FUNCTION "FRK_ModelRoot" : Int
{ S7_Optimized_Access := 'TRUE' }
VERSION : 0.1
VAR_INPUT
    Scope : String;
END_VAR
BEGIN
    #FRK_ModelRoot := 0;
    IF #Scope = 'StationA' THEN #FRK_ModelRoot := 1; RETURN; END_IF;
    IF #Scope = 'StationB' THEN #FRK_ModelRoot := 2; RETURN; END_IF;
END_FUNCTION
// Core model identities and cloned configuration are one owned catalog domain.
// Native UMAC/recipe CSV cannot replace its typed, root-scoped admission rules.
FUNCTION "FRK_ModelCodeValid" : Bool
{ S7_Optimized_Access := 'TRUE' }
VERSION : 0.1
VAR_INPUT Code : String; END_VAR
VAR_TEMP Index : Int; Value : Byte; END_VAR
BEGIN
    #FRK_ModelCodeValid := FALSE;
    IF LEN(#Code) < 1 OR LEN(#Code) > 64 THEN RETURN; END_IF;
    FOR #Index := 1 TO LEN(#Code) DO
        #Value := CHAR_TO_BYTE(#Code[#Index]);
        IF #Value < BYTE#32 OR #Value > BYTE#126 THEN RETURN; END_IF;
    END_FOR;
    #FRK_ModelCodeValid := TRUE;
END_FUNCTION

FUNCTION "FRK_ModelCrc" : DWord
{ S7_Optimized_Access := 'TRUE' }
VERSION : 0.1
VAR_IN_OUT Catalog : "FRK_ModelCatalog"; END_VAR
VAR_TEMP Work : DWord; Index : Int; Character : Int; Size : Int; Text : String[80]; END_VAR
BEGIN
    #Work := "FRK_CrcNumber"(Previous := DWORD#16#FFFFFFFF, Value := UINT_TO_UDINT(#Catalog.SchemaVersion));
    #Size := LEN(#Catalog.Scope);
    #Work := "FRK_CrcNumber"(Previous := #Work, Value := INT_TO_UDINT(#Size));
    FOR #Character := 1 TO #Size DO #Work := "FRK_CrcByte"(Previous := #Work, Value := CHAR_TO_BYTE(#Catalog.Scope[#Character])); END_FOR;
    #Work := "FRK_CrcNumber"(Previous := #Work, Value := INT_TO_UDINT(#Catalog.Capacity));
    #Work := "FRK_CrcNumber"(Previous := #Work, Value := INT_TO_UDINT(#Catalog.Count));
    #Work := "FRK_CrcNumber"(Previous := #Work, Value := #Catalog.Generation);
    FOR #Index := 1 TO 3 DO
        #Text := #Catalog.Codes[#Index]; #Size := LEN(#Text);
        #Work := "FRK_CrcNumber"(Previous := #Work, Value := INT_TO_UDINT(#Size));
        FOR #Character := 1 TO #Size DO #Work := "FRK_CrcByte"(Previous := #Work, Value := CHAR_TO_BYTE(#Text[#Character])); END_FOR;
    END_FOR;
    #FRK_ModelCrc := NOT #Work;
END_FUNCTION

FUNCTION "FRK_ModelValid" : Bool
{ S7_Optimized_Access := 'TRUE' }
VERSION : 0.1
VAR_INPUT RootIndex : Int; END_VAR
VAR_IN_OUT Catalog : "FRK_ModelCatalog"; END_VAR
VAR_TEMP Index : Int; Other : Int; END_VAR
BEGIN
    #FRK_ModelValid := FALSE;
    IF #RootIndex < 1 OR #RootIndex > 2 OR "FRK_ModelRoot"(Scope := #Catalog.Scope) <> #RootIndex THEN RETURN; END_IF;
    IF #Catalog.SchemaVersion <> 1 OR #Catalog.Generation = 0 OR #Catalog.Capacity <> 3
        OR #Catalog.Count < 2 OR #Catalog.Count > 3 THEN RETURN; END_IF;
    IF #Catalog.Codes[1] <> 'MODEL_A' OR #Catalog.Codes[2] <> 'MODEL_B' THEN RETURN; END_IF;
    FOR #Index := 1 TO #Catalog.Count DO
        IF NOT "FRK_ModelCodeValid"(Code := #Catalog.Codes[#Index]) THEN RETURN; END_IF;
        FOR #Other := 1 TO #Index - 1 DO
            IF #Catalog.Codes[#Index] = #Catalog.Codes[#Other] THEN RETURN; END_IF;
        END_FOR;
    END_FOR;
    FOR #Index := #Catalog.Count + 1 TO 3 DO
        IF #Catalog.Codes[#Index] <> '' THEN RETURN; END_IF;
    END_FOR;
    #FRK_ModelValid := #Catalog.Checksum = "FRK_ModelCrc"(Catalog := #Catalog);
END_FUNCTION

FUNCTION "FRK_ModelVirgin" : Bool
{ S7_Optimized_Access := 'TRUE' }
VERSION : 0.1
VAR_IN_OUT Catalog : "FRK_ModelCatalog"; END_VAR
VAR_TEMP Index : Int; END_VAR
BEGIN
    #FRK_ModelVirgin := FALSE;
    IF #Catalog.SchemaVersion <> 0 OR #Catalog.Scope <> '' OR #Catalog.Capacity <> 0 OR #Catalog.Count <> 0
        OR #Catalog.Generation <> 0 OR #Catalog.Checksum <> DWORD#0 THEN RETURN; END_IF;
    FOR #Index := 1 TO 3 DO IF #Catalog.Codes[#Index] <> '' THEN RETURN; END_IF; END_FOR;
    #FRK_ModelVirgin := TRUE;
END_FUNCTION

FUNCTION "FRK_ModelKnown" : Bool
{ S7_Optimized_Access := 'TRUE' }
VERSION : 0.1
VAR_INPUT RootIndex : Int; Code : String; END_VAR
VAR_TEMP Index : Int; END_VAR
BEGIN
    #FRK_ModelKnown := FALSE;
    IF #RootIndex < 1 OR #RootIndex > 2 OR #Code = '' THEN RETURN; END_IF;
    IF "FRK_ModelStore".Rows[#RootIndex].Count < 2 OR "FRK_ModelStore".Rows[#RootIndex].Count > 3 THEN RETURN; END_IF;
    FOR #Index := 1 TO "FRK_ModelStore".Rows[#RootIndex].Count DO
        IF "FRK_ModelStore".Rows[#RootIndex].Codes[#Index] = #Code THEN #FRK_ModelKnown := TRUE; RETURN; END_IF;
    END_FOR;
END_FUNCTION
FUNCTION "FRK_ModelCapture_R1" : Bool
{ S7_Optimized_Access := 'TRUE' }
VERSION : 0.1
VAR_IN_OUT
    Catalog : "FRK_ModelCatalog";
    Image : "FRK_ModelImage";
END_VAR
VAR_TEMP
    Index : Int;
    ModelSlot : Int;
    RowIndex : Int;
    Stored : Int;
END_VAR
BEGIN
    #FRK_ModelCapture_R1 := FALSE;
    IF NOT "FRK_ModelValid"(RootIndex := 1, Catalog := #Catalog) THEN RETURN; END_IF;
    #Image.Catalog := #Catalog; #Image.RecordCount := 0;
    FOR #Index := 1 TO 26 DO #Image.Rows[#Index] := "FRK_ModelRuntime".BlankSlot; END_FOR;
    FOR #ModelSlot := 3 TO #Catalog.Count DO
        #RowIndex := (#ModelSlot - 3) * 26 + 1;
        "FRK_CfgDef_DeclarationUnit"(FieldIndex := 1);
        #Stored := "FRK_ConfigFind"(Scope := 'StationA', Key := 'timeout', ModelCode := #Catalog.Codes[#ModelSlot]);
        IF #Stored = 0 OR NOT "FRK_ConfigGet"(Scope := 'StationA', ModelCode := #Catalog.Codes[#ModelSlot]) THEN RETURN; END_IF;
        #Image.Rows[#RowIndex] := "FRK_ConfigStore".Rows[#Stored];
        #Image.RecordCount := #Image.RecordCount + 1;
        #RowIndex := (#ModelSlot - 3) * 26 + 2;
        "FRK_CfgDef_DeclarationUnit"(FieldIndex := 2);
        #Stored := "FRK_ConfigFind"(Scope := 'StationA', Key := 'preset', ModelCode := #Catalog.Codes[#ModelSlot]);
        IF #Stored = 0 OR NOT "FRK_ConfigGet"(Scope := 'StationA', ModelCode := #Catalog.Codes[#ModelSlot]) THEN RETURN; END_IF;
        #Image.Rows[#RowIndex] := "FRK_ConfigStore".Rows[#Stored];
        #Image.RecordCount := #Image.RecordCount + 1;
        #RowIndex := (#ModelSlot - 3) * 26 + 3;
        "FRK_CfgDef_DeclarationUnit"(FieldIndex := 8);
        #Stored := "FRK_ConfigFind"(Scope := 'StationA', Key := 'idealCycleMs', ModelCode := #Catalog.Codes[#ModelSlot]);
        IF #Stored = 0 OR NOT "FRK_ConfigGet"(Scope := 'StationA', ModelCode := #Catalog.Codes[#ModelSlot]) THEN RETURN; END_IF;
        #Image.Rows[#RowIndex] := "FRK_ConfigStore".Rows[#Stored];
        #Image.RecordCount := #Image.RecordCount + 1;
        #RowIndex := (#ModelSlot - 3) * 26 + 4;
        "FRK_CfgDef_DeclarationUnit"(FieldIndex := 9);
        #Stored := "FRK_ConfigFind"(Scope := 'StationA', Key := 'baselineMs', ModelCode := #Catalog.Codes[#ModelSlot]);
        IF #Stored = 0 OR NOT "FRK_ConfigGet"(Scope := 'StationA', ModelCode := #Catalog.Codes[#ModelSlot]) THEN RETURN; END_IF;
        #Image.Rows[#RowIndex] := "FRK_ConfigStore".Rows[#Stored];
        #Image.RecordCount := #Image.RecordCount + 1;
        #RowIndex := (#ModelSlot - 3) * 26 + 5;
        "FRK_CfgDef_DeclarationCell"(FieldIndex := 1);
        #Stored := "FRK_ConfigFind"(Scope := 'StationA.Cell', Key := 'timeout', ModelCode := #Catalog.Codes[#ModelSlot]);
        IF #Stored = 0 OR NOT "FRK_ConfigGet"(Scope := 'StationA.Cell', ModelCode := #Catalog.Codes[#ModelSlot]) THEN RETURN; END_IF;
        #Image.Rows[#RowIndex] := "FRK_ConfigStore".Rows[#Stored];
        #Image.RecordCount := #Image.RecordCount + 1;
        #RowIndex := (#ModelSlot - 3) * 26 + 6;
        "FRK_CfgDef_DeclarationCell"(FieldIndex := 2);
        #Stored := "FRK_ConfigFind"(Scope := 'StationA.Cell', Key := 'preset', ModelCode := #Catalog.Codes[#ModelSlot]);
        IF #Stored = 0 OR NOT "FRK_ConfigGet"(Scope := 'StationA.Cell', ModelCode := #Catalog.Codes[#ModelSlot]) THEN RETURN; END_IF;
        #Image.Rows[#RowIndex] := "FRK_ConfigStore".Rows[#Stored];
        #Image.RecordCount := #Image.RecordCount + 1;
        #RowIndex := (#ModelSlot - 3) * 26 + 7;
        "FRK_CfgDef_DeclarationCylinder"(FieldIndex := 1);
        #Stored := "FRK_ConfigFind"(Scope := 'StationA.Cell.Clamp', Key := 'timeout', ModelCode := #Catalog.Codes[#ModelSlot]);
        IF #Stored = 0 OR NOT "FRK_ConfigGet"(Scope := 'StationA.Cell.Clamp', ModelCode := #Catalog.Codes[#ModelSlot]) THEN RETURN; END_IF;
        #Image.Rows[#RowIndex] := "FRK_ConfigStore".Rows[#Stored];
        #Image.RecordCount := #Image.RecordCount + 1;
        #RowIndex := (#ModelSlot - 3) * 26 + 8;
        "FRK_CfgDef_DeclarationCylinder"(FieldIndex := 2);
        #Stored := "FRK_ConfigFind"(Scope := 'StationA.Cell.Clamp', Key := 'preset', ModelCode := #Catalog.Codes[#ModelSlot]);
        IF #Stored = 0 OR NOT "FRK_ConfigGet"(Scope := 'StationA.Cell.Clamp', ModelCode := #Catalog.Codes[#ModelSlot]) THEN RETURN; END_IF;
        #Image.Rows[#RowIndex] := "FRK_ConfigStore".Rows[#Stored];
        #Image.RecordCount := #Image.RecordCount + 1;
        #RowIndex := (#ModelSlot - 3) * 26 + 9;
        "FRK_CfgDef_DeclarationCylinder"(FieldIndex := 1);
        #Stored := "FRK_ConfigFind"(Scope := 'StationA.Cell.Gate', Key := 'timeout', ModelCode := #Catalog.Codes[#ModelSlot]);
        IF #Stored = 0 OR NOT "FRK_ConfigGet"(Scope := 'StationA.Cell.Gate', ModelCode := #Catalog.Codes[#ModelSlot]) THEN RETURN; END_IF;
        #Image.Rows[#RowIndex] := "FRK_ConfigStore".Rows[#Stored];
        #Image.RecordCount := #Image.RecordCount + 1;
        #RowIndex := (#ModelSlot - 3) * 26 + 10;
        "FRK_CfgDef_DeclarationCylinder"(FieldIndex := 2);
        #Stored := "FRK_ConfigFind"(Scope := 'StationA.Cell.Gate', Key := 'preset', ModelCode := #Catalog.Codes[#ModelSlot]);
        IF #Stored = 0 OR NOT "FRK_ConfigGet"(Scope := 'StationA.Cell.Gate', ModelCode := #Catalog.Codes[#ModelSlot]) THEN RETURN; END_IF;
        #Image.Rows[#RowIndex] := "FRK_ConfigStore".Rows[#Stored];
        #Image.RecordCount := #Image.RecordCount + 1;
        #RowIndex := (#ModelSlot - 3) * 26 + 11;
        "FRK_CfgDef_SatelliteUnit"(FieldIndex := 1);
        #Stored := "FRK_ConfigFind"(Scope := 'StationA.Satellite', Key := 'timeout', ModelCode := #Catalog.Codes[#ModelSlot]);
        IF #Stored = 0 OR NOT "FRK_ConfigGet"(Scope := 'StationA.Satellite', ModelCode := #Catalog.Codes[#ModelSlot]) THEN RETURN; END_IF;
        #Image.Rows[#RowIndex] := "FRK_ConfigStore".Rows[#Stored];
        #Image.RecordCount := #Image.RecordCount + 1;
        #RowIndex := (#ModelSlot - 3) * 26 + 12;
        "FRK_CfgDef_SatelliteUnit"(FieldIndex := 2);
        #Stored := "FRK_ConfigFind"(Scope := 'StationA.Satellite', Key := 'preset', ModelCode := #Catalog.Codes[#ModelSlot]);
        IF #Stored = 0 OR NOT "FRK_ConfigGet"(Scope := 'StationA.Satellite', ModelCode := #Catalog.Codes[#ModelSlot]) THEN RETURN; END_IF;
        #Image.Rows[#RowIndex] := "FRK_ConfigStore".Rows[#Stored];
        #Image.RecordCount := #Image.RecordCount + 1;
        #RowIndex := (#ModelSlot - 3) * 26 + 13;
        "FRK_CfgDef_DeclarationCell"(FieldIndex := 1);
        #Stored := "FRK_ConfigFind"(Scope := 'StationA.Satellite.Cell', Key := 'timeout', ModelCode := #Catalog.Codes[#ModelSlot]);
        IF #Stored = 0 OR NOT "FRK_ConfigGet"(Scope := 'StationA.Satellite.Cell', ModelCode := #Catalog.Codes[#ModelSlot]) THEN RETURN; END_IF;
        #Image.Rows[#RowIndex] := "FRK_ConfigStore".Rows[#Stored];
        #Image.RecordCount := #Image.RecordCount + 1;
        #RowIndex := (#ModelSlot - 3) * 26 + 14;
        "FRK_CfgDef_DeclarationCell"(FieldIndex := 2);
        #Stored := "FRK_ConfigFind"(Scope := 'StationA.Satellite.Cell', Key := 'preset', ModelCode := #Catalog.Codes[#ModelSlot]);
        IF #Stored = 0 OR NOT "FRK_ConfigGet"(Scope := 'StationA.Satellite.Cell', ModelCode := #Catalog.Codes[#ModelSlot]) THEN RETURN; END_IF;
        #Image.Rows[#RowIndex] := "FRK_ConfigStore".Rows[#Stored];
        #Image.RecordCount := #Image.RecordCount + 1;
        #RowIndex := (#ModelSlot - 3) * 26 + 15;
        "FRK_CfgDef_DeclarationCylinder"(FieldIndex := 1);
        #Stored := "FRK_ConfigFind"(Scope := 'StationA.Satellite.Cell.Clamp', Key := 'timeout', ModelCode := #Catalog.Codes[#ModelSlot]);
        IF #Stored = 0 OR NOT "FRK_ConfigGet"(Scope := 'StationA.Satellite.Cell.Clamp', ModelCode := #Catalog.Codes[#ModelSlot]) THEN RETURN; END_IF;
        #Image.Rows[#RowIndex] := "FRK_ConfigStore".Rows[#Stored];
        #Image.RecordCount := #Image.RecordCount + 1;
        #RowIndex := (#ModelSlot - 3) * 26 + 16;
        "FRK_CfgDef_DeclarationCylinder"(FieldIndex := 2);
        #Stored := "FRK_ConfigFind"(Scope := 'StationA.Satellite.Cell.Clamp', Key := 'preset', ModelCode := #Catalog.Codes[#ModelSlot]);
        IF #Stored = 0 OR NOT "FRK_ConfigGet"(Scope := 'StationA.Satellite.Cell.Clamp', ModelCode := #Catalog.Codes[#ModelSlot]) THEN RETURN; END_IF;
        #Image.Rows[#RowIndex] := "FRK_ConfigStore".Rows[#Stored];
        #Image.RecordCount := #Image.RecordCount + 1;
        #RowIndex := (#ModelSlot - 3) * 26 + 17;
        "FRK_CfgDef_DeclarationCylinder"(FieldIndex := 1);
        #Stored := "FRK_ConfigFind"(Scope := 'StationA.Satellite.Cell.Gate', Key := 'timeout', ModelCode := #Catalog.Codes[#ModelSlot]);
        IF #Stored = 0 OR NOT "FRK_ConfigGet"(Scope := 'StationA.Satellite.Cell.Gate', ModelCode := #Catalog.Codes[#ModelSlot]) THEN RETURN; END_IF;
        #Image.Rows[#RowIndex] := "FRK_ConfigStore".Rows[#Stored];
        #Image.RecordCount := #Image.RecordCount + 1;
        #RowIndex := (#ModelSlot - 3) * 26 + 18;
        "FRK_CfgDef_DeclarationCylinder"(FieldIndex := 2);
        #Stored := "FRK_ConfigFind"(Scope := 'StationA.Satellite.Cell.Gate', Key := 'preset', ModelCode := #Catalog.Codes[#ModelSlot]);
        IF #Stored = 0 OR NOT "FRK_ConfigGet"(Scope := 'StationA.Satellite.Cell.Gate', ModelCode := #Catalog.Codes[#ModelSlot]) THEN RETURN; END_IF;
        #Image.Rows[#RowIndex] := "FRK_ConfigStore".Rows[#Stored];
        #Image.RecordCount := #Image.RecordCount + 1;
        #RowIndex := (#ModelSlot - 3) * 26 + 19;
        "FRK_CfgDef_InnerUnit"(FieldIndex := 1);
        #Stored := "FRK_ConfigFind"(Scope := 'StationA.Satellite.Inner', Key := 'timeout', ModelCode := #Catalog.Codes[#ModelSlot]);
        IF #Stored = 0 OR NOT "FRK_ConfigGet"(Scope := 'StationA.Satellite.Inner', ModelCode := #Catalog.Codes[#ModelSlot]) THEN RETURN; END_IF;
        #Image.Rows[#RowIndex] := "FRK_ConfigStore".Rows[#Stored];
        #Image.RecordCount := #Image.RecordCount + 1;
        #RowIndex := (#ModelSlot - 3) * 26 + 20;
        "FRK_CfgDef_InnerUnit"(FieldIndex := 2);
        #Stored := "FRK_ConfigFind"(Scope := 'StationA.Satellite.Inner', Key := 'preset', ModelCode := #Catalog.Codes[#ModelSlot]);
        IF #Stored = 0 OR NOT "FRK_ConfigGet"(Scope := 'StationA.Satellite.Inner', ModelCode := #Catalog.Codes[#ModelSlot]) THEN RETURN; END_IF;
        #Image.Rows[#RowIndex] := "FRK_ConfigStore".Rows[#Stored];
        #Image.RecordCount := #Image.RecordCount + 1;
        #RowIndex := (#ModelSlot - 3) * 26 + 21;
        "FRK_CfgDef_DeclarationCell"(FieldIndex := 1);
        #Stored := "FRK_ConfigFind"(Scope := 'StationA.Satellite.Inner.Cell', Key := 'timeout', ModelCode := #Catalog.Codes[#ModelSlot]);
        IF #Stored = 0 OR NOT "FRK_ConfigGet"(Scope := 'StationA.Satellite.Inner.Cell', ModelCode := #Catalog.Codes[#ModelSlot]) THEN RETURN; END_IF;
        #Image.Rows[#RowIndex] := "FRK_ConfigStore".Rows[#Stored];
        #Image.RecordCount := #Image.RecordCount + 1;
        #RowIndex := (#ModelSlot - 3) * 26 + 22;
        "FRK_CfgDef_DeclarationCell"(FieldIndex := 2);
        #Stored := "FRK_ConfigFind"(Scope := 'StationA.Satellite.Inner.Cell', Key := 'preset', ModelCode := #Catalog.Codes[#ModelSlot]);
        IF #Stored = 0 OR NOT "FRK_ConfigGet"(Scope := 'StationA.Satellite.Inner.Cell', ModelCode := #Catalog.Codes[#ModelSlot]) THEN RETURN; END_IF;
        #Image.Rows[#RowIndex] := "FRK_ConfigStore".Rows[#Stored];
        #Image.RecordCount := #Image.RecordCount + 1;
        #RowIndex := (#ModelSlot - 3) * 26 + 23;
        "FRK_CfgDef_DeclarationCylinder"(FieldIndex := 1);
        #Stored := "FRK_ConfigFind"(Scope := 'StationA.Satellite.Inner.Cell.Clamp', Key := 'timeout', ModelCode := #Catalog.Codes[#ModelSlot]);
        IF #Stored = 0 OR NOT "FRK_ConfigGet"(Scope := 'StationA.Satellite.Inner.Cell.Clamp', ModelCode := #Catalog.Codes[#ModelSlot]) THEN RETURN; END_IF;
        #Image.Rows[#RowIndex] := "FRK_ConfigStore".Rows[#Stored];
        #Image.RecordCount := #Image.RecordCount + 1;
        #RowIndex := (#ModelSlot - 3) * 26 + 24;
        "FRK_CfgDef_DeclarationCylinder"(FieldIndex := 2);
        #Stored := "FRK_ConfigFind"(Scope := 'StationA.Satellite.Inner.Cell.Clamp', Key := 'preset', ModelCode := #Catalog.Codes[#ModelSlot]);
        IF #Stored = 0 OR NOT "FRK_ConfigGet"(Scope := 'StationA.Satellite.Inner.Cell.Clamp', ModelCode := #Catalog.Codes[#ModelSlot]) THEN RETURN; END_IF;
        #Image.Rows[#RowIndex] := "FRK_ConfigStore".Rows[#Stored];
        #Image.RecordCount := #Image.RecordCount + 1;
        #RowIndex := (#ModelSlot - 3) * 26 + 25;
        "FRK_CfgDef_DeclarationCylinder"(FieldIndex := 1);
        #Stored := "FRK_ConfigFind"(Scope := 'StationA.Satellite.Inner.Cell.Gate', Key := 'timeout', ModelCode := #Catalog.Codes[#ModelSlot]);
        IF #Stored = 0 OR NOT "FRK_ConfigGet"(Scope := 'StationA.Satellite.Inner.Cell.Gate', ModelCode := #Catalog.Codes[#ModelSlot]) THEN RETURN; END_IF;
        #Image.Rows[#RowIndex] := "FRK_ConfigStore".Rows[#Stored];
        #Image.RecordCount := #Image.RecordCount + 1;
        #RowIndex := (#ModelSlot - 3) * 26 + 26;
        "FRK_CfgDef_DeclarationCylinder"(FieldIndex := 2);
        #Stored := "FRK_ConfigFind"(Scope := 'StationA.Satellite.Inner.Cell.Gate', Key := 'preset', ModelCode := #Catalog.Codes[#ModelSlot]);
        IF #Stored = 0 OR NOT "FRK_ConfigGet"(Scope := 'StationA.Satellite.Inner.Cell.Gate', ModelCode := #Catalog.Codes[#ModelSlot]) THEN RETURN; END_IF;
        #Image.Rows[#RowIndex] := "FRK_ConfigStore".Rows[#Stored];
        #Image.RecordCount := #Image.RecordCount + 1;
    END_FOR;
    #FRK_ModelCapture_R1 := TRUE;
END_FUNCTION
FUNCTION "FRK_ModelApply_R1" : Bool
{ S7_Optimized_Access := 'TRUE' }
VERSION : 0.1
VAR_IN_OUT
    Image : "FRK_ModelImage";
END_VAR
VAR_TEMP
    Index : Int;
    ModelSlot : Int;
    RowIndex : Int;
    Stored : Int;
    Targets : Array[1..32] of Int;
END_VAR
BEGIN
    #FRK_ModelApply_R1 := FALSE;
    IF NOT "FRK_ModelValid"(RootIndex := 1, Catalog := #Image.Catalog) THEN RETURN; END_IF;
    IF #Image.RecordCount <> (#Image.Catalog.Count - 2) * 26 THEN RETURN; END_IF;
    FOR #Index := 1 TO 32 DO #Targets[#Index] := 0; END_FOR;
    FOR #ModelSlot := 3 TO #Image.Catalog.Count DO
        #RowIndex := (#ModelSlot - 3) * 26 + 1;
        "FRK_CfgDef_DeclarationUnit"(FieldIndex := 1);
        IF NOT #Image.Rows[#RowIndex].Used OR #Image.Rows[#RowIndex].SchemaVersion <> "FRK_ConfigScratch".Schema
            OR #Image.Rows[#RowIndex].ModelCode <> #Image.Catalog.Codes[#ModelSlot]
            THEN RETURN; END_IF;
        IF NOT "FRK_ConfigRecordValid"(Scope := 'StationA', Record := #Image.Rows[#RowIndex].Record) THEN RETURN; END_IF;
        #Stored := "FRK_ConfigReserve"(Scope := 'StationA', Key := 'timeout', ModelCode := #Image.Catalog.Codes[#ModelSlot], Reserved := #Targets);
        IF #Stored < 1 OR #Stored > 212 THEN RETURN; END_IF;
        #Targets[#RowIndex] := #Stored;
        #RowIndex := (#ModelSlot - 3) * 26 + 2;
        "FRK_CfgDef_DeclarationUnit"(FieldIndex := 2);
        IF NOT #Image.Rows[#RowIndex].Used OR #Image.Rows[#RowIndex].SchemaVersion <> "FRK_ConfigScratch".Schema
            OR #Image.Rows[#RowIndex].ModelCode <> #Image.Catalog.Codes[#ModelSlot]
            THEN RETURN; END_IF;
        IF NOT "FRK_ConfigRecordValid"(Scope := 'StationA', Record := #Image.Rows[#RowIndex].Record) THEN RETURN; END_IF;
        #Stored := "FRK_ConfigReserve"(Scope := 'StationA', Key := 'preset', ModelCode := #Image.Catalog.Codes[#ModelSlot], Reserved := #Targets);
        IF #Stored < 1 OR #Stored > 212 THEN RETURN; END_IF;
        #Targets[#RowIndex] := #Stored;
        #RowIndex := (#ModelSlot - 3) * 26 + 3;
        "FRK_CfgDef_DeclarationUnit"(FieldIndex := 8);
        IF NOT #Image.Rows[#RowIndex].Used OR #Image.Rows[#RowIndex].SchemaVersion <> "FRK_ConfigScratch".Schema
            OR #Image.Rows[#RowIndex].ModelCode <> #Image.Catalog.Codes[#ModelSlot]
            THEN RETURN; END_IF;
        IF NOT "FRK_ConfigRecordValid"(Scope := 'StationA', Record := #Image.Rows[#RowIndex].Record) THEN RETURN; END_IF;
        #Stored := "FRK_ConfigReserve"(Scope := 'StationA', Key := 'idealCycleMs', ModelCode := #Image.Catalog.Codes[#ModelSlot], Reserved := #Targets);
        IF #Stored < 1 OR #Stored > 212 THEN RETURN; END_IF;
        #Targets[#RowIndex] := #Stored;
        #RowIndex := (#ModelSlot - 3) * 26 + 4;
        "FRK_CfgDef_DeclarationUnit"(FieldIndex := 9);
        IF NOT #Image.Rows[#RowIndex].Used OR #Image.Rows[#RowIndex].SchemaVersion <> "FRK_ConfigScratch".Schema
            OR #Image.Rows[#RowIndex].ModelCode <> #Image.Catalog.Codes[#ModelSlot]
            THEN RETURN; END_IF;
        IF NOT "FRK_ConfigRecordValid"(Scope := 'StationA', Record := #Image.Rows[#RowIndex].Record) THEN RETURN; END_IF;
        #Stored := "FRK_ConfigReserve"(Scope := 'StationA', Key := 'baselineMs', ModelCode := #Image.Catalog.Codes[#ModelSlot], Reserved := #Targets);
        IF #Stored < 1 OR #Stored > 212 THEN RETURN; END_IF;
        #Targets[#RowIndex] := #Stored;
        #RowIndex := (#ModelSlot - 3) * 26 + 5;
        "FRK_CfgDef_DeclarationCell"(FieldIndex := 1);
        IF NOT #Image.Rows[#RowIndex].Used OR #Image.Rows[#RowIndex].SchemaVersion <> "FRK_ConfigScratch".Schema
            OR #Image.Rows[#RowIndex].ModelCode <> #Image.Catalog.Codes[#ModelSlot]
            THEN RETURN; END_IF;
        IF NOT "FRK_ConfigRecordValid"(Scope := 'StationA.Cell', Record := #Image.Rows[#RowIndex].Record) THEN RETURN; END_IF;
        #Stored := "FRK_ConfigReserve"(Scope := 'StationA.Cell', Key := 'timeout', ModelCode := #Image.Catalog.Codes[#ModelSlot], Reserved := #Targets);
        IF #Stored < 1 OR #Stored > 212 THEN RETURN; END_IF;
        #Targets[#RowIndex] := #Stored;
        #RowIndex := (#ModelSlot - 3) * 26 + 6;
        "FRK_CfgDef_DeclarationCell"(FieldIndex := 2);
        IF NOT #Image.Rows[#RowIndex].Used OR #Image.Rows[#RowIndex].SchemaVersion <> "FRK_ConfigScratch".Schema
            OR #Image.Rows[#RowIndex].ModelCode <> #Image.Catalog.Codes[#ModelSlot]
            THEN RETURN; END_IF;
        IF NOT "FRK_ConfigRecordValid"(Scope := 'StationA.Cell', Record := #Image.Rows[#RowIndex].Record) THEN RETURN; END_IF;
        #Stored := "FRK_ConfigReserve"(Scope := 'StationA.Cell', Key := 'preset', ModelCode := #Image.Catalog.Codes[#ModelSlot], Reserved := #Targets);
        IF #Stored < 1 OR #Stored > 212 THEN RETURN; END_IF;
        #Targets[#RowIndex] := #Stored;
        #RowIndex := (#ModelSlot - 3) * 26 + 7;
        "FRK_CfgDef_DeclarationCylinder"(FieldIndex := 1);
        IF NOT #Image.Rows[#RowIndex].Used OR #Image.Rows[#RowIndex].SchemaVersion <> "FRK_ConfigScratch".Schema
            OR #Image.Rows[#RowIndex].ModelCode <> #Image.Catalog.Codes[#ModelSlot]
            THEN RETURN; END_IF;
        IF NOT "FRK_ConfigRecordValid"(Scope := 'StationA.Cell.Clamp', Record := #Image.Rows[#RowIndex].Record) THEN RETURN; END_IF;
        #Stored := "FRK_ConfigReserve"(Scope := 'StationA.Cell.Clamp', Key := 'timeout', ModelCode := #Image.Catalog.Codes[#ModelSlot], Reserved := #Targets);
        IF #Stored < 1 OR #Stored > 212 THEN RETURN; END_IF;
        #Targets[#RowIndex] := #Stored;
        #RowIndex := (#ModelSlot - 3) * 26 + 8;
        "FRK_CfgDef_DeclarationCylinder"(FieldIndex := 2);
        IF NOT #Image.Rows[#RowIndex].Used OR #Image.Rows[#RowIndex].SchemaVersion <> "FRK_ConfigScratch".Schema
            OR #Image.Rows[#RowIndex].ModelCode <> #Image.Catalog.Codes[#ModelSlot]
            THEN RETURN; END_IF;
        IF NOT "FRK_ConfigRecordValid"(Scope := 'StationA.Cell.Clamp', Record := #Image.Rows[#RowIndex].Record) THEN RETURN; END_IF;
        #Stored := "FRK_ConfigReserve"(Scope := 'StationA.Cell.Clamp', Key := 'preset', ModelCode := #Image.Catalog.Codes[#ModelSlot], Reserved := #Targets);
        IF #Stored < 1 OR #Stored > 212 THEN RETURN; END_IF;
        #Targets[#RowIndex] := #Stored;
        #RowIndex := (#ModelSlot - 3) * 26 + 9;
        "FRK_CfgDef_DeclarationCylinder"(FieldIndex := 1);
        IF NOT #Image.Rows[#RowIndex].Used OR #Image.Rows[#RowIndex].SchemaVersion <> "FRK_ConfigScratch".Schema
            OR #Image.Rows[#RowIndex].ModelCode <> #Image.Catalog.Codes[#ModelSlot]
            THEN RETURN; END_IF;
        IF NOT "FRK_ConfigRecordValid"(Scope := 'StationA.Cell.Gate', Record := #Image.Rows[#RowIndex].Record) THEN RETURN; END_IF;
        #Stored := "FRK_ConfigReserve"(Scope := 'StationA.Cell.Gate', Key := 'timeout', ModelCode := #Image.Catalog.Codes[#ModelSlot], Reserved := #Targets);
        IF #Stored < 1 OR #Stored > 212 THEN RETURN; END_IF;
        #Targets[#RowIndex] := #Stored;
        #RowIndex := (#ModelSlot - 3) * 26 + 10;
        "FRK_CfgDef_DeclarationCylinder"(FieldIndex := 2);
        IF NOT #Image.Rows[#RowIndex].Used OR #Image.Rows[#RowIndex].SchemaVersion <> "FRK_ConfigScratch".Schema
            OR #Image.Rows[#RowIndex].ModelCode <> #Image.Catalog.Codes[#ModelSlot]
            THEN RETURN; END_IF;
        IF NOT "FRK_ConfigRecordValid"(Scope := 'StationA.Cell.Gate', Record := #Image.Rows[#RowIndex].Record) THEN RETURN; END_IF;
        #Stored := "FRK_ConfigReserve"(Scope := 'StationA.Cell.Gate', Key := 'preset', ModelCode := #Image.Catalog.Codes[#ModelSlot], Reserved := #Targets);
        IF #Stored < 1 OR #Stored > 212 THEN RETURN; END_IF;
        #Targets[#RowIndex] := #Stored;
        #RowIndex := (#ModelSlot - 3) * 26 + 11;
        "FRK_CfgDef_SatelliteUnit"(FieldIndex := 1);
        IF NOT #Image.Rows[#RowIndex].Used OR #Image.Rows[#RowIndex].SchemaVersion <> "FRK_ConfigScratch".Schema
            OR #Image.Rows[#RowIndex].ModelCode <> #Image.Catalog.Codes[#ModelSlot]
            THEN RETURN; END_IF;
        IF NOT "FRK_ConfigRecordValid"(Scope := 'StationA.Satellite', Record := #Image.Rows[#RowIndex].Record) THEN RETURN; END_IF;
        #Stored := "FRK_ConfigReserve"(Scope := 'StationA.Satellite', Key := 'timeout', ModelCode := #Image.Catalog.Codes[#ModelSlot], Reserved := #Targets);
        IF #Stored < 1 OR #Stored > 212 THEN RETURN; END_IF;
        #Targets[#RowIndex] := #Stored;
        #RowIndex := (#ModelSlot - 3) * 26 + 12;
        "FRK_CfgDef_SatelliteUnit"(FieldIndex := 2);
        IF NOT #Image.Rows[#RowIndex].Used OR #Image.Rows[#RowIndex].SchemaVersion <> "FRK_ConfigScratch".Schema
            OR #Image.Rows[#RowIndex].ModelCode <> #Image.Catalog.Codes[#ModelSlot]
            THEN RETURN; END_IF;
        IF NOT "FRK_ConfigRecordValid"(Scope := 'StationA.Satellite', Record := #Image.Rows[#RowIndex].Record) THEN RETURN; END_IF;
        #Stored := "FRK_ConfigReserve"(Scope := 'StationA.Satellite', Key := 'preset', ModelCode := #Image.Catalog.Codes[#ModelSlot], Reserved := #Targets);
        IF #Stored < 1 OR #Stored > 212 THEN RETURN; END_IF;
        #Targets[#RowIndex] := #Stored;
        #RowIndex := (#ModelSlot - 3) * 26 + 13;
        "FRK_CfgDef_DeclarationCell"(FieldIndex := 1);
        IF NOT #Image.Rows[#RowIndex].Used OR #Image.Rows[#RowIndex].SchemaVersion <> "FRK_ConfigScratch".Schema
            OR #Image.Rows[#RowIndex].ModelCode <> #Image.Catalog.Codes[#ModelSlot]
            THEN RETURN; END_IF;
        IF NOT "FRK_ConfigRecordValid"(Scope := 'StationA.Satellite.Cell', Record := #Image.Rows[#RowIndex].Record) THEN RETURN; END_IF;
        #Stored := "FRK_ConfigReserve"(Scope := 'StationA.Satellite.Cell', Key := 'timeout', ModelCode := #Image.Catalog.Codes[#ModelSlot], Reserved := #Targets);
        IF #Stored < 1 OR #Stored > 212 THEN RETURN; END_IF;
        #Targets[#RowIndex] := #Stored;
        #RowIndex := (#ModelSlot - 3) * 26 + 14;
        "FRK_CfgDef_DeclarationCell"(FieldIndex := 2);
        IF NOT #Image.Rows[#RowIndex].Used OR #Image.Rows[#RowIndex].SchemaVersion <> "FRK_ConfigScratch".Schema
            OR #Image.Rows[#RowIndex].ModelCode <> #Image.Catalog.Codes[#ModelSlot]
            THEN RETURN; END_IF;
        IF NOT "FRK_ConfigRecordValid"(Scope := 'StationA.Satellite.Cell', Record := #Image.Rows[#RowIndex].Record) THEN RETURN; END_IF;
        #Stored := "FRK_ConfigReserve"(Scope := 'StationA.Satellite.Cell', Key := 'preset', ModelCode := #Image.Catalog.Codes[#ModelSlot], Reserved := #Targets);
        IF #Stored < 1 OR #Stored > 212 THEN RETURN; END_IF;
        #Targets[#RowIndex] := #Stored;
        #RowIndex := (#ModelSlot - 3) * 26 + 15;
        "FRK_CfgDef_DeclarationCylinder"(FieldIndex := 1);
        IF NOT #Image.Rows[#RowIndex].Used OR #Image.Rows[#RowIndex].SchemaVersion <> "FRK_ConfigScratch".Schema
            OR #Image.Rows[#RowIndex].ModelCode <> #Image.Catalog.Codes[#ModelSlot]
            THEN RETURN; END_IF;
        IF NOT "FRK_ConfigRecordValid"(Scope := 'StationA.Satellite.Cell.Clamp', Record := #Image.Rows[#RowIndex].Record) THEN RETURN; END_IF;
        #Stored := "FRK_ConfigReserve"(Scope := 'StationA.Satellite.Cell.Clamp', Key := 'timeout', ModelCode := #Image.Catalog.Codes[#ModelSlot], Reserved := #Targets);
        IF #Stored < 1 OR #Stored > 212 THEN RETURN; END_IF;
        #Targets[#RowIndex] := #Stored;
        #RowIndex := (#ModelSlot - 3) * 26 + 16;
        "FRK_CfgDef_DeclarationCylinder"(FieldIndex := 2);
        IF NOT #Image.Rows[#RowIndex].Used OR #Image.Rows[#RowIndex].SchemaVersion <> "FRK_ConfigScratch".Schema
            OR #Image.Rows[#RowIndex].ModelCode <> #Image.Catalog.Codes[#ModelSlot]
            THEN RETURN; END_IF;
        IF NOT "FRK_ConfigRecordValid"(Scope := 'StationA.Satellite.Cell.Clamp', Record := #Image.Rows[#RowIndex].Record) THEN RETURN; END_IF;
        #Stored := "FRK_ConfigReserve"(Scope := 'StationA.Satellite.Cell.Clamp', Key := 'preset', ModelCode := #Image.Catalog.Codes[#ModelSlot], Reserved := #Targets);
        IF #Stored < 1 OR #Stored > 212 THEN RETURN; END_IF;
        #Targets[#RowIndex] := #Stored;
        #RowIndex := (#ModelSlot - 3) * 26 + 17;
        "FRK_CfgDef_DeclarationCylinder"(FieldIndex := 1);
        IF NOT #Image.Rows[#RowIndex].Used OR #Image.Rows[#RowIndex].SchemaVersion <> "FRK_ConfigScratch".Schema
            OR #Image.Rows[#RowIndex].ModelCode <> #Image.Catalog.Codes[#ModelSlot]
            THEN RETURN; END_IF;
        IF NOT "FRK_ConfigRecordValid"(Scope := 'StationA.Satellite.Cell.Gate', Record := #Image.Rows[#RowIndex].Record) THEN RETURN; END_IF;
        #Stored := "FRK_ConfigReserve"(Scope := 'StationA.Satellite.Cell.Gate', Key := 'timeout', ModelCode := #Image.Catalog.Codes[#ModelSlot], Reserved := #Targets);
        IF #Stored < 1 OR #Stored > 212 THEN RETURN; END_IF;
        #Targets[#RowIndex] := #Stored;
        #RowIndex := (#ModelSlot - 3) * 26 + 18;
        "FRK_CfgDef_DeclarationCylinder"(FieldIndex := 2);
        IF NOT #Image.Rows[#RowIndex].Used OR #Image.Rows[#RowIndex].SchemaVersion <> "FRK_ConfigScratch".Schema
            OR #Image.Rows[#RowIndex].ModelCode <> #Image.Catalog.Codes[#ModelSlot]
            THEN RETURN; END_IF;
        IF NOT "FRK_ConfigRecordValid"(Scope := 'StationA.Satellite.Cell.Gate', Record := #Image.Rows[#RowIndex].Record) THEN RETURN; END_IF;
        #Stored := "FRK_ConfigReserve"(Scope := 'StationA.Satellite.Cell.Gate', Key := 'preset', ModelCode := #Image.Catalog.Codes[#ModelSlot], Reserved := #Targets);
        IF #Stored < 1 OR #Stored > 212 THEN RETURN; END_IF;
        #Targets[#RowIndex] := #Stored;
        #RowIndex := (#ModelSlot - 3) * 26 + 19;
        "FRK_CfgDef_InnerUnit"(FieldIndex := 1);
        IF NOT #Image.Rows[#RowIndex].Used OR #Image.Rows[#RowIndex].SchemaVersion <> "FRK_ConfigScratch".Schema
            OR #Image.Rows[#RowIndex].ModelCode <> #Image.Catalog.Codes[#ModelSlot]
            THEN RETURN; END_IF;
        IF NOT "FRK_ConfigRecordValid"(Scope := 'StationA.Satellite.Inner', Record := #Image.Rows[#RowIndex].Record) THEN RETURN; END_IF;
        #Stored := "FRK_ConfigReserve"(Scope := 'StationA.Satellite.Inner', Key := 'timeout', ModelCode := #Image.Catalog.Codes[#ModelSlot], Reserved := #Targets);
        IF #Stored < 1 OR #Stored > 212 THEN RETURN; END_IF;
        #Targets[#RowIndex] := #Stored;
        #RowIndex := (#ModelSlot - 3) * 26 + 20;
        "FRK_CfgDef_InnerUnit"(FieldIndex := 2);
        IF NOT #Image.Rows[#RowIndex].Used OR #Image.Rows[#RowIndex].SchemaVersion <> "FRK_ConfigScratch".Schema
            OR #Image.Rows[#RowIndex].ModelCode <> #Image.Catalog.Codes[#ModelSlot]
            THEN RETURN; END_IF;
        IF NOT "FRK_ConfigRecordValid"(Scope := 'StationA.Satellite.Inner', Record := #Image.Rows[#RowIndex].Record) THEN RETURN; END_IF;
        #Stored := "FRK_ConfigReserve"(Scope := 'StationA.Satellite.Inner', Key := 'preset', ModelCode := #Image.Catalog.Codes[#ModelSlot], Reserved := #Targets);
        IF #Stored < 1 OR #Stored > 212 THEN RETURN; END_IF;
        #Targets[#RowIndex] := #Stored;
        #RowIndex := (#ModelSlot - 3) * 26 + 21;
        "FRK_CfgDef_DeclarationCell"(FieldIndex := 1);
        IF NOT #Image.Rows[#RowIndex].Used OR #Image.Rows[#RowIndex].SchemaVersion <> "FRK_ConfigScratch".Schema
            OR #Image.Rows[#RowIndex].ModelCode <> #Image.Catalog.Codes[#ModelSlot]
            THEN RETURN; END_IF;
        IF NOT "FRK_ConfigRecordValid"(Scope := 'StationA.Satellite.Inner.Cell', Record := #Image.Rows[#RowIndex].Record) THEN RETURN; END_IF;
        #Stored := "FRK_ConfigReserve"(Scope := 'StationA.Satellite.Inner.Cell', Key := 'timeout', ModelCode := #Image.Catalog.Codes[#ModelSlot], Reserved := #Targets);
        IF #Stored < 1 OR #Stored > 212 THEN RETURN; END_IF;
        #Targets[#RowIndex] := #Stored;
        #RowIndex := (#ModelSlot - 3) * 26 + 22;
        "FRK_CfgDef_DeclarationCell"(FieldIndex := 2);
        IF NOT #Image.Rows[#RowIndex].Used OR #Image.Rows[#RowIndex].SchemaVersion <> "FRK_ConfigScratch".Schema
            OR #Image.Rows[#RowIndex].ModelCode <> #Image.Catalog.Codes[#ModelSlot]
            THEN RETURN; END_IF;
        IF NOT "FRK_ConfigRecordValid"(Scope := 'StationA.Satellite.Inner.Cell', Record := #Image.Rows[#RowIndex].Record) THEN RETURN; END_IF;
        #Stored := "FRK_ConfigReserve"(Scope := 'StationA.Satellite.Inner.Cell', Key := 'preset', ModelCode := #Image.Catalog.Codes[#ModelSlot], Reserved := #Targets);
        IF #Stored < 1 OR #Stored > 212 THEN RETURN; END_IF;
        #Targets[#RowIndex] := #Stored;
        #RowIndex := (#ModelSlot - 3) * 26 + 23;
        "FRK_CfgDef_DeclarationCylinder"(FieldIndex := 1);
        IF NOT #Image.Rows[#RowIndex].Used OR #Image.Rows[#RowIndex].SchemaVersion <> "FRK_ConfigScratch".Schema
            OR #Image.Rows[#RowIndex].ModelCode <> #Image.Catalog.Codes[#ModelSlot]
            THEN RETURN; END_IF;
        IF NOT "FRK_ConfigRecordValid"(Scope := 'StationA.Satellite.Inner.Cell.Clamp', Record := #Image.Rows[#RowIndex].Record) THEN RETURN; END_IF;
        #Stored := "FRK_ConfigReserve"(Scope := 'StationA.Satellite.Inner.Cell.Clamp', Key := 'timeout', ModelCode := #Image.Catalog.Codes[#ModelSlot], Reserved := #Targets);
        IF #Stored < 1 OR #Stored > 212 THEN RETURN; END_IF;
        #Targets[#RowIndex] := #Stored;
        #RowIndex := (#ModelSlot - 3) * 26 + 24;
        "FRK_CfgDef_DeclarationCylinder"(FieldIndex := 2);
        IF NOT #Image.Rows[#RowIndex].Used OR #Image.Rows[#RowIndex].SchemaVersion <> "FRK_ConfigScratch".Schema
            OR #Image.Rows[#RowIndex].ModelCode <> #Image.Catalog.Codes[#ModelSlot]
            THEN RETURN; END_IF;
        IF NOT "FRK_ConfigRecordValid"(Scope := 'StationA.Satellite.Inner.Cell.Clamp', Record := #Image.Rows[#RowIndex].Record) THEN RETURN; END_IF;
        #Stored := "FRK_ConfigReserve"(Scope := 'StationA.Satellite.Inner.Cell.Clamp', Key := 'preset', ModelCode := #Image.Catalog.Codes[#ModelSlot], Reserved := #Targets);
        IF #Stored < 1 OR #Stored > 212 THEN RETURN; END_IF;
        #Targets[#RowIndex] := #Stored;
        #RowIndex := (#ModelSlot - 3) * 26 + 25;
        "FRK_CfgDef_DeclarationCylinder"(FieldIndex := 1);
        IF NOT #Image.Rows[#RowIndex].Used OR #Image.Rows[#RowIndex].SchemaVersion <> "FRK_ConfigScratch".Schema
            OR #Image.Rows[#RowIndex].ModelCode <> #Image.Catalog.Codes[#ModelSlot]
            THEN RETURN; END_IF;
        IF NOT "FRK_ConfigRecordValid"(Scope := 'StationA.Satellite.Inner.Cell.Gate', Record := #Image.Rows[#RowIndex].Record) THEN RETURN; END_IF;
        #Stored := "FRK_ConfigReserve"(Scope := 'StationA.Satellite.Inner.Cell.Gate', Key := 'timeout', ModelCode := #Image.Catalog.Codes[#ModelSlot], Reserved := #Targets);
        IF #Stored < 1 OR #Stored > 212 THEN RETURN; END_IF;
        #Targets[#RowIndex] := #Stored;
        #RowIndex := (#ModelSlot - 3) * 26 + 26;
        "FRK_CfgDef_DeclarationCylinder"(FieldIndex := 2);
        IF NOT #Image.Rows[#RowIndex].Used OR #Image.Rows[#RowIndex].SchemaVersion <> "FRK_ConfigScratch".Schema
            OR #Image.Rows[#RowIndex].ModelCode <> #Image.Catalog.Codes[#ModelSlot]
            THEN RETURN; END_IF;
        IF NOT "FRK_ConfigRecordValid"(Scope := 'StationA.Satellite.Inner.Cell.Gate', Record := #Image.Rows[#RowIndex].Record) THEN RETURN; END_IF;
        #Stored := "FRK_ConfigReserve"(Scope := 'StationA.Satellite.Inner.Cell.Gate', Key := 'preset', ModelCode := #Image.Catalog.Codes[#ModelSlot], Reserved := #Targets);
        IF #Stored < 1 OR #Stored > 212 THEN RETURN; END_IF;
        #Targets[#RowIndex] := #Stored;
    END_FOR;
    FOR #Index := 1 TO #Image.RecordCount DO
        "FRK_ConfigStore".Rows[#Targets[#Index]] := #Image.Rows[#Index];
    END_FOR;
    "FRK_ModelStore".Rows[1] := #Image.Catalog;
    "FRK_ConfigStore".SchemaVersion := 1;
    #FRK_ModelApply_R1 := TRUE;
END_FUNCTION
FUNCTION "FRK_ModelCapture_R2" : Bool
{ S7_Optimized_Access := 'TRUE' }
VERSION : 0.1
VAR_IN_OUT
    Catalog : "FRK_ModelCatalog";
    Image : "FRK_ModelImage";
END_VAR
VAR_TEMP
    Index : Int;
    ModelSlot : Int;
    RowIndex : Int;
    Stored : Int;
END_VAR
BEGIN
    #FRK_ModelCapture_R2 := FALSE;
    IF NOT "FRK_ModelValid"(RootIndex := 2, Catalog := #Catalog) THEN RETURN; END_IF;
    #Image.Catalog := #Catalog; #Image.RecordCount := 0;
    FOR #Index := 1 TO 26 DO #Image.Rows[#Index] := "FRK_ModelRuntime".BlankSlot; END_FOR;
    FOR #ModelSlot := 3 TO #Catalog.Count DO
        #RowIndex := (#ModelSlot - 3) * 26 + 1;
        "FRK_CfgDef_DeclarationUnit"(FieldIndex := 1);
        #Stored := "FRK_ConfigFind"(Scope := 'StationB', Key := 'timeout', ModelCode := #Catalog.Codes[#ModelSlot]);
        IF #Stored = 0 OR NOT "FRK_ConfigGet"(Scope := 'StationB', ModelCode := #Catalog.Codes[#ModelSlot]) THEN RETURN; END_IF;
        #Image.Rows[#RowIndex] := "FRK_ConfigStore".Rows[#Stored];
        #Image.RecordCount := #Image.RecordCount + 1;
        #RowIndex := (#ModelSlot - 3) * 26 + 2;
        "FRK_CfgDef_DeclarationUnit"(FieldIndex := 2);
        #Stored := "FRK_ConfigFind"(Scope := 'StationB', Key := 'preset', ModelCode := #Catalog.Codes[#ModelSlot]);
        IF #Stored = 0 OR NOT "FRK_ConfigGet"(Scope := 'StationB', ModelCode := #Catalog.Codes[#ModelSlot]) THEN RETURN; END_IF;
        #Image.Rows[#RowIndex] := "FRK_ConfigStore".Rows[#Stored];
        #Image.RecordCount := #Image.RecordCount + 1;
        #RowIndex := (#ModelSlot - 3) * 26 + 3;
        "FRK_CfgDef_DeclarationUnit"(FieldIndex := 8);
        #Stored := "FRK_ConfigFind"(Scope := 'StationB', Key := 'idealCycleMs', ModelCode := #Catalog.Codes[#ModelSlot]);
        IF #Stored = 0 OR NOT "FRK_ConfigGet"(Scope := 'StationB', ModelCode := #Catalog.Codes[#ModelSlot]) THEN RETURN; END_IF;
        #Image.Rows[#RowIndex] := "FRK_ConfigStore".Rows[#Stored];
        #Image.RecordCount := #Image.RecordCount + 1;
        #RowIndex := (#ModelSlot - 3) * 26 + 4;
        "FRK_CfgDef_DeclarationUnit"(FieldIndex := 9);
        #Stored := "FRK_ConfigFind"(Scope := 'StationB', Key := 'baselineMs', ModelCode := #Catalog.Codes[#ModelSlot]);
        IF #Stored = 0 OR NOT "FRK_ConfigGet"(Scope := 'StationB', ModelCode := #Catalog.Codes[#ModelSlot]) THEN RETURN; END_IF;
        #Image.Rows[#RowIndex] := "FRK_ConfigStore".Rows[#Stored];
        #Image.RecordCount := #Image.RecordCount + 1;
        #RowIndex := (#ModelSlot - 3) * 26 + 5;
        "FRK_CfgDef_DeclarationCell"(FieldIndex := 1);
        #Stored := "FRK_ConfigFind"(Scope := 'StationB.Cell', Key := 'timeout', ModelCode := #Catalog.Codes[#ModelSlot]);
        IF #Stored = 0 OR NOT "FRK_ConfigGet"(Scope := 'StationB.Cell', ModelCode := #Catalog.Codes[#ModelSlot]) THEN RETURN; END_IF;
        #Image.Rows[#RowIndex] := "FRK_ConfigStore".Rows[#Stored];
        #Image.RecordCount := #Image.RecordCount + 1;
        #RowIndex := (#ModelSlot - 3) * 26 + 6;
        "FRK_CfgDef_DeclarationCell"(FieldIndex := 2);
        #Stored := "FRK_ConfigFind"(Scope := 'StationB.Cell', Key := 'preset', ModelCode := #Catalog.Codes[#ModelSlot]);
        IF #Stored = 0 OR NOT "FRK_ConfigGet"(Scope := 'StationB.Cell', ModelCode := #Catalog.Codes[#ModelSlot]) THEN RETURN; END_IF;
        #Image.Rows[#RowIndex] := "FRK_ConfigStore".Rows[#Stored];
        #Image.RecordCount := #Image.RecordCount + 1;
        #RowIndex := (#ModelSlot - 3) * 26 + 7;
        "FRK_CfgDef_DeclarationCylinder"(FieldIndex := 1);
        #Stored := "FRK_ConfigFind"(Scope := 'StationB.Cell.Clamp', Key := 'timeout', ModelCode := #Catalog.Codes[#ModelSlot]);
        IF #Stored = 0 OR NOT "FRK_ConfigGet"(Scope := 'StationB.Cell.Clamp', ModelCode := #Catalog.Codes[#ModelSlot]) THEN RETURN; END_IF;
        #Image.Rows[#RowIndex] := "FRK_ConfigStore".Rows[#Stored];
        #Image.RecordCount := #Image.RecordCount + 1;
        #RowIndex := (#ModelSlot - 3) * 26 + 8;
        "FRK_CfgDef_DeclarationCylinder"(FieldIndex := 2);
        #Stored := "FRK_ConfigFind"(Scope := 'StationB.Cell.Clamp', Key := 'preset', ModelCode := #Catalog.Codes[#ModelSlot]);
        IF #Stored = 0 OR NOT "FRK_ConfigGet"(Scope := 'StationB.Cell.Clamp', ModelCode := #Catalog.Codes[#ModelSlot]) THEN RETURN; END_IF;
        #Image.Rows[#RowIndex] := "FRK_ConfigStore".Rows[#Stored];
        #Image.RecordCount := #Image.RecordCount + 1;
        #RowIndex := (#ModelSlot - 3) * 26 + 9;
        "FRK_CfgDef_DeclarationCylinder"(FieldIndex := 1);
        #Stored := "FRK_ConfigFind"(Scope := 'StationB.Cell.Gate', Key := 'timeout', ModelCode := #Catalog.Codes[#ModelSlot]);
        IF #Stored = 0 OR NOT "FRK_ConfigGet"(Scope := 'StationB.Cell.Gate', ModelCode := #Catalog.Codes[#ModelSlot]) THEN RETURN; END_IF;
        #Image.Rows[#RowIndex] := "FRK_ConfigStore".Rows[#Stored];
        #Image.RecordCount := #Image.RecordCount + 1;
        #RowIndex := (#ModelSlot - 3) * 26 + 10;
        "FRK_CfgDef_DeclarationCylinder"(FieldIndex := 2);
        #Stored := "FRK_ConfigFind"(Scope := 'StationB.Cell.Gate', Key := 'preset', ModelCode := #Catalog.Codes[#ModelSlot]);
        IF #Stored = 0 OR NOT "FRK_ConfigGet"(Scope := 'StationB.Cell.Gate', ModelCode := #Catalog.Codes[#ModelSlot]) THEN RETURN; END_IF;
        #Image.Rows[#RowIndex] := "FRK_ConfigStore".Rows[#Stored];
        #Image.RecordCount := #Image.RecordCount + 1;
        #RowIndex := (#ModelSlot - 3) * 26 + 11;
        "FRK_CfgDef_SatelliteUnit"(FieldIndex := 1);
        #Stored := "FRK_ConfigFind"(Scope := 'StationB.Satellite', Key := 'timeout', ModelCode := #Catalog.Codes[#ModelSlot]);
        IF #Stored = 0 OR NOT "FRK_ConfigGet"(Scope := 'StationB.Satellite', ModelCode := #Catalog.Codes[#ModelSlot]) THEN RETURN; END_IF;
        #Image.Rows[#RowIndex] := "FRK_ConfigStore".Rows[#Stored];
        #Image.RecordCount := #Image.RecordCount + 1;
        #RowIndex := (#ModelSlot - 3) * 26 + 12;
        "FRK_CfgDef_SatelliteUnit"(FieldIndex := 2);
        #Stored := "FRK_ConfigFind"(Scope := 'StationB.Satellite', Key := 'preset', ModelCode := #Catalog.Codes[#ModelSlot]);
        IF #Stored = 0 OR NOT "FRK_ConfigGet"(Scope := 'StationB.Satellite', ModelCode := #Catalog.Codes[#ModelSlot]) THEN RETURN; END_IF;
        #Image.Rows[#RowIndex] := "FRK_ConfigStore".Rows[#Stored];
        #Image.RecordCount := #Image.RecordCount + 1;
        #RowIndex := (#ModelSlot - 3) * 26 + 13;
        "FRK_CfgDef_DeclarationCell"(FieldIndex := 1);
        #Stored := "FRK_ConfigFind"(Scope := 'StationB.Satellite.Cell', Key := 'timeout', ModelCode := #Catalog.Codes[#ModelSlot]);
        IF #Stored = 0 OR NOT "FRK_ConfigGet"(Scope := 'StationB.Satellite.Cell', ModelCode := #Catalog.Codes[#ModelSlot]) THEN RETURN; END_IF;
        #Image.Rows[#RowIndex] := "FRK_ConfigStore".Rows[#Stored];
        #Image.RecordCount := #Image.RecordCount + 1;
        #RowIndex := (#ModelSlot - 3) * 26 + 14;
        "FRK_CfgDef_DeclarationCell"(FieldIndex := 2);
        #Stored := "FRK_ConfigFind"(Scope := 'StationB.Satellite.Cell', Key := 'preset', ModelCode := #Catalog.Codes[#ModelSlot]);
        IF #Stored = 0 OR NOT "FRK_ConfigGet"(Scope := 'StationB.Satellite.Cell', ModelCode := #Catalog.Codes[#ModelSlot]) THEN RETURN; END_IF;
        #Image.Rows[#RowIndex] := "FRK_ConfigStore".Rows[#Stored];
        #Image.RecordCount := #Image.RecordCount + 1;
        #RowIndex := (#ModelSlot - 3) * 26 + 15;
        "FRK_CfgDef_DeclarationCylinder"(FieldIndex := 1);
        #Stored := "FRK_ConfigFind"(Scope := 'StationB.Satellite.Cell.Clamp', Key := 'timeout', ModelCode := #Catalog.Codes[#ModelSlot]);
        IF #Stored = 0 OR NOT "FRK_ConfigGet"(Scope := 'StationB.Satellite.Cell.Clamp', ModelCode := #Catalog.Codes[#ModelSlot]) THEN RETURN; END_IF;
        #Image.Rows[#RowIndex] := "FRK_ConfigStore".Rows[#Stored];
        #Image.RecordCount := #Image.RecordCount + 1;
        #RowIndex := (#ModelSlot - 3) * 26 + 16;
        "FRK_CfgDef_DeclarationCylinder"(FieldIndex := 2);
        #Stored := "FRK_ConfigFind"(Scope := 'StationB.Satellite.Cell.Clamp', Key := 'preset', ModelCode := #Catalog.Codes[#ModelSlot]);
        IF #Stored = 0 OR NOT "FRK_ConfigGet"(Scope := 'StationB.Satellite.Cell.Clamp', ModelCode := #Catalog.Codes[#ModelSlot]) THEN RETURN; END_IF;
        #Image.Rows[#RowIndex] := "FRK_ConfigStore".Rows[#Stored];
        #Image.RecordCount := #Image.RecordCount + 1;
        #RowIndex := (#ModelSlot - 3) * 26 + 17;
        "FRK_CfgDef_DeclarationCylinder"(FieldIndex := 1);
        #Stored := "FRK_ConfigFind"(Scope := 'StationB.Satellite.Cell.Gate', Key := 'timeout', ModelCode := #Catalog.Codes[#ModelSlot]);
        IF #Stored = 0 OR NOT "FRK_ConfigGet"(Scope := 'StationB.Satellite.Cell.Gate', ModelCode := #Catalog.Codes[#ModelSlot]) THEN RETURN; END_IF;
        #Image.Rows[#RowIndex] := "FRK_ConfigStore".Rows[#Stored];
        #Image.RecordCount := #Image.RecordCount + 1;
        #RowIndex := (#ModelSlot - 3) * 26 + 18;
        "FRK_CfgDef_DeclarationCylinder"(FieldIndex := 2);
        #Stored := "FRK_ConfigFind"(Scope := 'StationB.Satellite.Cell.Gate', Key := 'preset', ModelCode := #Catalog.Codes[#ModelSlot]);
        IF #Stored = 0 OR NOT "FRK_ConfigGet"(Scope := 'StationB.Satellite.Cell.Gate', ModelCode := #Catalog.Codes[#ModelSlot]) THEN RETURN; END_IF;
        #Image.Rows[#RowIndex] := "FRK_ConfigStore".Rows[#Stored];
        #Image.RecordCount := #Image.RecordCount + 1;
        #RowIndex := (#ModelSlot - 3) * 26 + 19;
        "FRK_CfgDef_InnerUnit"(FieldIndex := 1);
        #Stored := "FRK_ConfigFind"(Scope := 'StationB.Satellite.Inner', Key := 'timeout', ModelCode := #Catalog.Codes[#ModelSlot]);
        IF #Stored = 0 OR NOT "FRK_ConfigGet"(Scope := 'StationB.Satellite.Inner', ModelCode := #Catalog.Codes[#ModelSlot]) THEN RETURN; END_IF;
        #Image.Rows[#RowIndex] := "FRK_ConfigStore".Rows[#Stored];
        #Image.RecordCount := #Image.RecordCount + 1;
        #RowIndex := (#ModelSlot - 3) * 26 + 20;
        "FRK_CfgDef_InnerUnit"(FieldIndex := 2);
        #Stored := "FRK_ConfigFind"(Scope := 'StationB.Satellite.Inner', Key := 'preset', ModelCode := #Catalog.Codes[#ModelSlot]);
        IF #Stored = 0 OR NOT "FRK_ConfigGet"(Scope := 'StationB.Satellite.Inner', ModelCode := #Catalog.Codes[#ModelSlot]) THEN RETURN; END_IF;
        #Image.Rows[#RowIndex] := "FRK_ConfigStore".Rows[#Stored];
        #Image.RecordCount := #Image.RecordCount + 1;
        #RowIndex := (#ModelSlot - 3) * 26 + 21;
        "FRK_CfgDef_DeclarationCell"(FieldIndex := 1);
        #Stored := "FRK_ConfigFind"(Scope := 'StationB.Satellite.Inner.Cell', Key := 'timeout', ModelCode := #Catalog.Codes[#ModelSlot]);
        IF #Stored = 0 OR NOT "FRK_ConfigGet"(Scope := 'StationB.Satellite.Inner.Cell', ModelCode := #Catalog.Codes[#ModelSlot]) THEN RETURN; END_IF;
        #Image.Rows[#RowIndex] := "FRK_ConfigStore".Rows[#Stored];
        #Image.RecordCount := #Image.RecordCount + 1;
        #RowIndex := (#ModelSlot - 3) * 26 + 22;
        "FRK_CfgDef_DeclarationCell"(FieldIndex := 2);
        #Stored := "FRK_ConfigFind"(Scope := 'StationB.Satellite.Inner.Cell', Key := 'preset', ModelCode := #Catalog.Codes[#ModelSlot]);
        IF #Stored = 0 OR NOT "FRK_ConfigGet"(Scope := 'StationB.Satellite.Inner.Cell', ModelCode := #Catalog.Codes[#ModelSlot]) THEN RETURN; END_IF;
        #Image.Rows[#RowIndex] := "FRK_ConfigStore".Rows[#Stored];
        #Image.RecordCount := #Image.RecordCount + 1;
        #RowIndex := (#ModelSlot - 3) * 26 + 23;
        "FRK_CfgDef_DeclarationCylinder"(FieldIndex := 1);
        #Stored := "FRK_ConfigFind"(Scope := 'StationB.Satellite.Inner.Cell.Clamp', Key := 'timeout', ModelCode := #Catalog.Codes[#ModelSlot]);
        IF #Stored = 0 OR NOT "FRK_ConfigGet"(Scope := 'StationB.Satellite.Inner.Cell.Clamp', ModelCode := #Catalog.Codes[#ModelSlot]) THEN RETURN; END_IF;
        #Image.Rows[#RowIndex] := "FRK_ConfigStore".Rows[#Stored];
        #Image.RecordCount := #Image.RecordCount + 1;
        #RowIndex := (#ModelSlot - 3) * 26 + 24;
        "FRK_CfgDef_DeclarationCylinder"(FieldIndex := 2);
        #Stored := "FRK_ConfigFind"(Scope := 'StationB.Satellite.Inner.Cell.Clamp', Key := 'preset', ModelCode := #Catalog.Codes[#ModelSlot]);
        IF #Stored = 0 OR NOT "FRK_ConfigGet"(Scope := 'StationB.Satellite.Inner.Cell.Clamp', ModelCode := #Catalog.Codes[#ModelSlot]) THEN RETURN; END_IF;
        #Image.Rows[#RowIndex] := "FRK_ConfigStore".Rows[#Stored];
        #Image.RecordCount := #Image.RecordCount + 1;
        #RowIndex := (#ModelSlot - 3) * 26 + 25;
        "FRK_CfgDef_DeclarationCylinder"(FieldIndex := 1);
        #Stored := "FRK_ConfigFind"(Scope := 'StationB.Satellite.Inner.Cell.Gate', Key := 'timeout', ModelCode := #Catalog.Codes[#ModelSlot]);
        IF #Stored = 0 OR NOT "FRK_ConfigGet"(Scope := 'StationB.Satellite.Inner.Cell.Gate', ModelCode := #Catalog.Codes[#ModelSlot]) THEN RETURN; END_IF;
        #Image.Rows[#RowIndex] := "FRK_ConfigStore".Rows[#Stored];
        #Image.RecordCount := #Image.RecordCount + 1;
        #RowIndex := (#ModelSlot - 3) * 26 + 26;
        "FRK_CfgDef_DeclarationCylinder"(FieldIndex := 2);
        #Stored := "FRK_ConfigFind"(Scope := 'StationB.Satellite.Inner.Cell.Gate', Key := 'preset', ModelCode := #Catalog.Codes[#ModelSlot]);
        IF #Stored = 0 OR NOT "FRK_ConfigGet"(Scope := 'StationB.Satellite.Inner.Cell.Gate', ModelCode := #Catalog.Codes[#ModelSlot]) THEN RETURN; END_IF;
        #Image.Rows[#RowIndex] := "FRK_ConfigStore".Rows[#Stored];
        #Image.RecordCount := #Image.RecordCount + 1;
    END_FOR;
    #FRK_ModelCapture_R2 := TRUE;
END_FUNCTION
FUNCTION "FRK_ModelApply_R2" : Bool
{ S7_Optimized_Access := 'TRUE' }
VERSION : 0.1
VAR_IN_OUT
    Image : "FRK_ModelImage";
END_VAR
VAR_TEMP
    Index : Int;
    ModelSlot : Int;
    RowIndex : Int;
    Stored : Int;
    Targets : Array[1..32] of Int;
END_VAR
BEGIN
    #FRK_ModelApply_R2 := FALSE;
    IF NOT "FRK_ModelValid"(RootIndex := 2, Catalog := #Image.Catalog) THEN RETURN; END_IF;
    IF #Image.RecordCount <> (#Image.Catalog.Count - 2) * 26 THEN RETURN; END_IF;
    FOR #Index := 1 TO 32 DO #Targets[#Index] := 0; END_FOR;
    FOR #ModelSlot := 3 TO #Image.Catalog.Count DO
        #RowIndex := (#ModelSlot - 3) * 26 + 1;
        "FRK_CfgDef_DeclarationUnit"(FieldIndex := 1);
        IF NOT #Image.Rows[#RowIndex].Used OR #Image.Rows[#RowIndex].SchemaVersion <> "FRK_ConfigScratch".Schema
            OR #Image.Rows[#RowIndex].ModelCode <> #Image.Catalog.Codes[#ModelSlot]
            THEN RETURN; END_IF;
        IF NOT "FRK_ConfigRecordValid"(Scope := 'StationB', Record := #Image.Rows[#RowIndex].Record) THEN RETURN; END_IF;
        #Stored := "FRK_ConfigReserve"(Scope := 'StationB', Key := 'timeout', ModelCode := #Image.Catalog.Codes[#ModelSlot], Reserved := #Targets);
        IF #Stored < 1 OR #Stored > 212 THEN RETURN; END_IF;
        #Targets[#RowIndex] := #Stored;
        #RowIndex := (#ModelSlot - 3) * 26 + 2;
        "FRK_CfgDef_DeclarationUnit"(FieldIndex := 2);
        IF NOT #Image.Rows[#RowIndex].Used OR #Image.Rows[#RowIndex].SchemaVersion <> "FRK_ConfigScratch".Schema
            OR #Image.Rows[#RowIndex].ModelCode <> #Image.Catalog.Codes[#ModelSlot]
            THEN RETURN; END_IF;
        IF NOT "FRK_ConfigRecordValid"(Scope := 'StationB', Record := #Image.Rows[#RowIndex].Record) THEN RETURN; END_IF;
        #Stored := "FRK_ConfigReserve"(Scope := 'StationB', Key := 'preset', ModelCode := #Image.Catalog.Codes[#ModelSlot], Reserved := #Targets);
        IF #Stored < 1 OR #Stored > 212 THEN RETURN; END_IF;
        #Targets[#RowIndex] := #Stored;
        #RowIndex := (#ModelSlot - 3) * 26 + 3;
        "FRK_CfgDef_DeclarationUnit"(FieldIndex := 8);
        IF NOT #Image.Rows[#RowIndex].Used OR #Image.Rows[#RowIndex].SchemaVersion <> "FRK_ConfigScratch".Schema
            OR #Image.Rows[#RowIndex].ModelCode <> #Image.Catalog.Codes[#ModelSlot]
            THEN RETURN; END_IF;
        IF NOT "FRK_ConfigRecordValid"(Scope := 'StationB', Record := #Image.Rows[#RowIndex].Record) THEN RETURN; END_IF;
        #Stored := "FRK_ConfigReserve"(Scope := 'StationB', Key := 'idealCycleMs', ModelCode := #Image.Catalog.Codes[#ModelSlot], Reserved := #Targets);
        IF #Stored < 1 OR #Stored > 212 THEN RETURN; END_IF;
        #Targets[#RowIndex] := #Stored;
        #RowIndex := (#ModelSlot - 3) * 26 + 4;
        "FRK_CfgDef_DeclarationUnit"(FieldIndex := 9);
        IF NOT #Image.Rows[#RowIndex].Used OR #Image.Rows[#RowIndex].SchemaVersion <> "FRK_ConfigScratch".Schema
            OR #Image.Rows[#RowIndex].ModelCode <> #Image.Catalog.Codes[#ModelSlot]
            THEN RETURN; END_IF;
        IF NOT "FRK_ConfigRecordValid"(Scope := 'StationB', Record := #Image.Rows[#RowIndex].Record) THEN RETURN; END_IF;
        #Stored := "FRK_ConfigReserve"(Scope := 'StationB', Key := 'baselineMs', ModelCode := #Image.Catalog.Codes[#ModelSlot], Reserved := #Targets);
        IF #Stored < 1 OR #Stored > 212 THEN RETURN; END_IF;
        #Targets[#RowIndex] := #Stored;
        #RowIndex := (#ModelSlot - 3) * 26 + 5;
        "FRK_CfgDef_DeclarationCell"(FieldIndex := 1);
        IF NOT #Image.Rows[#RowIndex].Used OR #Image.Rows[#RowIndex].SchemaVersion <> "FRK_ConfigScratch".Schema
            OR #Image.Rows[#RowIndex].ModelCode <> #Image.Catalog.Codes[#ModelSlot]
            THEN RETURN; END_IF;
        IF NOT "FRK_ConfigRecordValid"(Scope := 'StationB.Cell', Record := #Image.Rows[#RowIndex].Record) THEN RETURN; END_IF;
        #Stored := "FRK_ConfigReserve"(Scope := 'StationB.Cell', Key := 'timeout', ModelCode := #Image.Catalog.Codes[#ModelSlot], Reserved := #Targets);
        IF #Stored < 1 OR #Stored > 212 THEN RETURN; END_IF;
        #Targets[#RowIndex] := #Stored;
        #RowIndex := (#ModelSlot - 3) * 26 + 6;
        "FRK_CfgDef_DeclarationCell"(FieldIndex := 2);
        IF NOT #Image.Rows[#RowIndex].Used OR #Image.Rows[#RowIndex].SchemaVersion <> "FRK_ConfigScratch".Schema
            OR #Image.Rows[#RowIndex].ModelCode <> #Image.Catalog.Codes[#ModelSlot]
            THEN RETURN; END_IF;
        IF NOT "FRK_ConfigRecordValid"(Scope := 'StationB.Cell', Record := #Image.Rows[#RowIndex].Record) THEN RETURN; END_IF;
        #Stored := "FRK_ConfigReserve"(Scope := 'StationB.Cell', Key := 'preset', ModelCode := #Image.Catalog.Codes[#ModelSlot], Reserved := #Targets);
        IF #Stored < 1 OR #Stored > 212 THEN RETURN; END_IF;
        #Targets[#RowIndex] := #Stored;
        #RowIndex := (#ModelSlot - 3) * 26 + 7;
        "FRK_CfgDef_DeclarationCylinder"(FieldIndex := 1);
        IF NOT #Image.Rows[#RowIndex].Used OR #Image.Rows[#RowIndex].SchemaVersion <> "FRK_ConfigScratch".Schema
            OR #Image.Rows[#RowIndex].ModelCode <> #Image.Catalog.Codes[#ModelSlot]
            THEN RETURN; END_IF;
        IF NOT "FRK_ConfigRecordValid"(Scope := 'StationB.Cell.Clamp', Record := #Image.Rows[#RowIndex].Record) THEN RETURN; END_IF;
        #Stored := "FRK_ConfigReserve"(Scope := 'StationB.Cell.Clamp', Key := 'timeout', ModelCode := #Image.Catalog.Codes[#ModelSlot], Reserved := #Targets);
        IF #Stored < 1 OR #Stored > 212 THEN RETURN; END_IF;
        #Targets[#RowIndex] := #Stored;
        #RowIndex := (#ModelSlot - 3) * 26 + 8;
        "FRK_CfgDef_DeclarationCylinder"(FieldIndex := 2);
        IF NOT #Image.Rows[#RowIndex].Used OR #Image.Rows[#RowIndex].SchemaVersion <> "FRK_ConfigScratch".Schema
            OR #Image.Rows[#RowIndex].ModelCode <> #Image.Catalog.Codes[#ModelSlot]
            THEN RETURN; END_IF;
        IF NOT "FRK_ConfigRecordValid"(Scope := 'StationB.Cell.Clamp', Record := #Image.Rows[#RowIndex].Record) THEN RETURN; END_IF;
        #Stored := "FRK_ConfigReserve"(Scope := 'StationB.Cell.Clamp', Key := 'preset', ModelCode := #Image.Catalog.Codes[#ModelSlot], Reserved := #Targets);
        IF #Stored < 1 OR #Stored > 212 THEN RETURN; END_IF;
        #Targets[#RowIndex] := #Stored;
        #RowIndex := (#ModelSlot - 3) * 26 + 9;
        "FRK_CfgDef_DeclarationCylinder"(FieldIndex := 1);
        IF NOT #Image.Rows[#RowIndex].Used OR #Image.Rows[#RowIndex].SchemaVersion <> "FRK_ConfigScratch".Schema
            OR #Image.Rows[#RowIndex].ModelCode <> #Image.Catalog.Codes[#ModelSlot]
            THEN RETURN; END_IF;
        IF NOT "FRK_ConfigRecordValid"(Scope := 'StationB.Cell.Gate', Record := #Image.Rows[#RowIndex].Record) THEN RETURN; END_IF;
        #Stored := "FRK_ConfigReserve"(Scope := 'StationB.Cell.Gate', Key := 'timeout', ModelCode := #Image.Catalog.Codes[#ModelSlot], Reserved := #Targets);
        IF #Stored < 1 OR #Stored > 212 THEN RETURN; END_IF;
        #Targets[#RowIndex] := #Stored;
        #RowIndex := (#ModelSlot - 3) * 26 + 10;
        "FRK_CfgDef_DeclarationCylinder"(FieldIndex := 2);
        IF NOT #Image.Rows[#RowIndex].Used OR #Image.Rows[#RowIndex].SchemaVersion <> "FRK_ConfigScratch".Schema
            OR #Image.Rows[#RowIndex].ModelCode <> #Image.Catalog.Codes[#ModelSlot]
            THEN RETURN; END_IF;
        IF NOT "FRK_ConfigRecordValid"(Scope := 'StationB.Cell.Gate', Record := #Image.Rows[#RowIndex].Record) THEN RETURN; END_IF;
        #Stored := "FRK_ConfigReserve"(Scope := 'StationB.Cell.Gate', Key := 'preset', ModelCode := #Image.Catalog.Codes[#ModelSlot], Reserved := #Targets);
        IF #Stored < 1 OR #Stored > 212 THEN RETURN; END_IF;
        #Targets[#RowIndex] := #Stored;
        #RowIndex := (#ModelSlot - 3) * 26 + 11;
        "FRK_CfgDef_SatelliteUnit"(FieldIndex := 1);
        IF NOT #Image.Rows[#RowIndex].Used OR #Image.Rows[#RowIndex].SchemaVersion <> "FRK_ConfigScratch".Schema
            OR #Image.Rows[#RowIndex].ModelCode <> #Image.Catalog.Codes[#ModelSlot]
            THEN RETURN; END_IF;
        IF NOT "FRK_ConfigRecordValid"(Scope := 'StationB.Satellite', Record := #Image.Rows[#RowIndex].Record) THEN RETURN; END_IF;
        #Stored := "FRK_ConfigReserve"(Scope := 'StationB.Satellite', Key := 'timeout', ModelCode := #Image.Catalog.Codes[#ModelSlot], Reserved := #Targets);
        IF #Stored < 1 OR #Stored > 212 THEN RETURN; END_IF;
        #Targets[#RowIndex] := #Stored;
        #RowIndex := (#ModelSlot - 3) * 26 + 12;
        "FRK_CfgDef_SatelliteUnit"(FieldIndex := 2);
        IF NOT #Image.Rows[#RowIndex].Used OR #Image.Rows[#RowIndex].SchemaVersion <> "FRK_ConfigScratch".Schema
            OR #Image.Rows[#RowIndex].ModelCode <> #Image.Catalog.Codes[#ModelSlot]
            THEN RETURN; END_IF;
        IF NOT "FRK_ConfigRecordValid"(Scope := 'StationB.Satellite', Record := #Image.Rows[#RowIndex].Record) THEN RETURN; END_IF;
        #Stored := "FRK_ConfigReserve"(Scope := 'StationB.Satellite', Key := 'preset', ModelCode := #Image.Catalog.Codes[#ModelSlot], Reserved := #Targets);
        IF #Stored < 1 OR #Stored > 212 THEN RETURN; END_IF;
        #Targets[#RowIndex] := #Stored;
        #RowIndex := (#ModelSlot - 3) * 26 + 13;
        "FRK_CfgDef_DeclarationCell"(FieldIndex := 1);
        IF NOT #Image.Rows[#RowIndex].Used OR #Image.Rows[#RowIndex].SchemaVersion <> "FRK_ConfigScratch".Schema
            OR #Image.Rows[#RowIndex].ModelCode <> #Image.Catalog.Codes[#ModelSlot]
            THEN RETURN; END_IF;
        IF NOT "FRK_ConfigRecordValid"(Scope := 'StationB.Satellite.Cell', Record := #Image.Rows[#RowIndex].Record) THEN RETURN; END_IF;
        #Stored := "FRK_ConfigReserve"(Scope := 'StationB.Satellite.Cell', Key := 'timeout', ModelCode := #Image.Catalog.Codes[#ModelSlot], Reserved := #Targets);
        IF #Stored < 1 OR #Stored > 212 THEN RETURN; END_IF;
        #Targets[#RowIndex] := #Stored;
        #RowIndex := (#ModelSlot - 3) * 26 + 14;
        "FRK_CfgDef_DeclarationCell"(FieldIndex := 2);
        IF NOT #Image.Rows[#RowIndex].Used OR #Image.Rows[#RowIndex].SchemaVersion <> "FRK_ConfigScratch".Schema
            OR #Image.Rows[#RowIndex].ModelCode <> #Image.Catalog.Codes[#ModelSlot]
            THEN RETURN; END_IF;
        IF NOT "FRK_ConfigRecordValid"(Scope := 'StationB.Satellite.Cell', Record := #Image.Rows[#RowIndex].Record) THEN RETURN; END_IF;
        #Stored := "FRK_ConfigReserve"(Scope := 'StationB.Satellite.Cell', Key := 'preset', ModelCode := #Image.Catalog.Codes[#ModelSlot], Reserved := #Targets);
        IF #Stored < 1 OR #Stored > 212 THEN RETURN; END_IF;
        #Targets[#RowIndex] := #Stored;
        #RowIndex := (#ModelSlot - 3) * 26 + 15;
        "FRK_CfgDef_DeclarationCylinder"(FieldIndex := 1);
        IF NOT #Image.Rows[#RowIndex].Used OR #Image.Rows[#RowIndex].SchemaVersion <> "FRK_ConfigScratch".Schema
            OR #Image.Rows[#RowIndex].ModelCode <> #Image.Catalog.Codes[#ModelSlot]
            THEN RETURN; END_IF;
        IF NOT "FRK_ConfigRecordValid"(Scope := 'StationB.Satellite.Cell.Clamp', Record := #Image.Rows[#RowIndex].Record) THEN RETURN; END_IF;
        #Stored := "FRK_ConfigReserve"(Scope := 'StationB.Satellite.Cell.Clamp', Key := 'timeout', ModelCode := #Image.Catalog.Codes[#ModelSlot], Reserved := #Targets);
        IF #Stored < 1 OR #Stored > 212 THEN RETURN; END_IF;
        #Targets[#RowIndex] := #Stored;
        #RowIndex := (#ModelSlot - 3) * 26 + 16;
        "FRK_CfgDef_DeclarationCylinder"(FieldIndex := 2);
        IF NOT #Image.Rows[#RowIndex].Used OR #Image.Rows[#RowIndex].SchemaVersion <> "FRK_ConfigScratch".Schema
            OR #Image.Rows[#RowIndex].ModelCode <> #Image.Catalog.Codes[#ModelSlot]
            THEN RETURN; END_IF;
        IF NOT "FRK_ConfigRecordValid"(Scope := 'StationB.Satellite.Cell.Clamp', Record := #Image.Rows[#RowIndex].Record) THEN RETURN; END_IF;
        #Stored := "FRK_ConfigReserve"(Scope := 'StationB.Satellite.Cell.Clamp', Key := 'preset', ModelCode := #Image.Catalog.Codes[#ModelSlot], Reserved := #Targets);
        IF #Stored < 1 OR #Stored > 212 THEN RETURN; END_IF;
        #Targets[#RowIndex] := #Stored;
        #RowIndex := (#ModelSlot - 3) * 26 + 17;
        "FRK_CfgDef_DeclarationCylinder"(FieldIndex := 1);
        IF NOT #Image.Rows[#RowIndex].Used OR #Image.Rows[#RowIndex].SchemaVersion <> "FRK_ConfigScratch".Schema
            OR #Image.Rows[#RowIndex].ModelCode <> #Image.Catalog.Codes[#ModelSlot]
            THEN RETURN; END_IF;
        IF NOT "FRK_ConfigRecordValid"(Scope := 'StationB.Satellite.Cell.Gate', Record := #Image.Rows[#RowIndex].Record) THEN RETURN; END_IF;
        #Stored := "FRK_ConfigReserve"(Scope := 'StationB.Satellite.Cell.Gate', Key := 'timeout', ModelCode := #Image.Catalog.Codes[#ModelSlot], Reserved := #Targets);
        IF #Stored < 1 OR #Stored > 212 THEN RETURN; END_IF;
        #Targets[#RowIndex] := #Stored;
        #RowIndex := (#ModelSlot - 3) * 26 + 18;
        "FRK_CfgDef_DeclarationCylinder"(FieldIndex := 2);
        IF NOT #Image.Rows[#RowIndex].Used OR #Image.Rows[#RowIndex].SchemaVersion <> "FRK_ConfigScratch".Schema
            OR #Image.Rows[#RowIndex].ModelCode <> #Image.Catalog.Codes[#ModelSlot]
            THEN RETURN; END_IF;
        IF NOT "FRK_ConfigRecordValid"(Scope := 'StationB.Satellite.Cell.Gate', Record := #Image.Rows[#RowIndex].Record) THEN RETURN; END_IF;
        #Stored := "FRK_ConfigReserve"(Scope := 'StationB.Satellite.Cell.Gate', Key := 'preset', ModelCode := #Image.Catalog.Codes[#ModelSlot], Reserved := #Targets);
        IF #Stored < 1 OR #Stored > 212 THEN RETURN; END_IF;
        #Targets[#RowIndex] := #Stored;
        #RowIndex := (#ModelSlot - 3) * 26 + 19;
        "FRK_CfgDef_InnerUnit"(FieldIndex := 1);
        IF NOT #Image.Rows[#RowIndex].Used OR #Image.Rows[#RowIndex].SchemaVersion <> "FRK_ConfigScratch".Schema
            OR #Image.Rows[#RowIndex].ModelCode <> #Image.Catalog.Codes[#ModelSlot]
            THEN RETURN; END_IF;
        IF NOT "FRK_ConfigRecordValid"(Scope := 'StationB.Satellite.Inner', Record := #Image.Rows[#RowIndex].Record) THEN RETURN; END_IF;
        #Stored := "FRK_ConfigReserve"(Scope := 'StationB.Satellite.Inner', Key := 'timeout', ModelCode := #Image.Catalog.Codes[#ModelSlot], Reserved := #Targets);
        IF #Stored < 1 OR #Stored > 212 THEN RETURN; END_IF;
        #Targets[#RowIndex] := #Stored;
        #RowIndex := (#ModelSlot - 3) * 26 + 20;
        "FRK_CfgDef_InnerUnit"(FieldIndex := 2);
        IF NOT #Image.Rows[#RowIndex].Used OR #Image.Rows[#RowIndex].SchemaVersion <> "FRK_ConfigScratch".Schema
            OR #Image.Rows[#RowIndex].ModelCode <> #Image.Catalog.Codes[#ModelSlot]
            THEN RETURN; END_IF;
        IF NOT "FRK_ConfigRecordValid"(Scope := 'StationB.Satellite.Inner', Record := #Image.Rows[#RowIndex].Record) THEN RETURN; END_IF;
        #Stored := "FRK_ConfigReserve"(Scope := 'StationB.Satellite.Inner', Key := 'preset', ModelCode := #Image.Catalog.Codes[#ModelSlot], Reserved := #Targets);
        IF #Stored < 1 OR #Stored > 212 THEN RETURN; END_IF;
        #Targets[#RowIndex] := #Stored;
        #RowIndex := (#ModelSlot - 3) * 26 + 21;
        "FRK_CfgDef_DeclarationCell"(FieldIndex := 1);
        IF NOT #Image.Rows[#RowIndex].Used OR #Image.Rows[#RowIndex].SchemaVersion <> "FRK_ConfigScratch".Schema
            OR #Image.Rows[#RowIndex].ModelCode <> #Image.Catalog.Codes[#ModelSlot]
            THEN RETURN; END_IF;
        IF NOT "FRK_ConfigRecordValid"(Scope := 'StationB.Satellite.Inner.Cell', Record := #Image.Rows[#RowIndex].Record) THEN RETURN; END_IF;
        #Stored := "FRK_ConfigReserve"(Scope := 'StationB.Satellite.Inner.Cell', Key := 'timeout', ModelCode := #Image.Catalog.Codes[#ModelSlot], Reserved := #Targets);
        IF #Stored < 1 OR #Stored > 212 THEN RETURN; END_IF;
        #Targets[#RowIndex] := #Stored;
        #RowIndex := (#ModelSlot - 3) * 26 + 22;
        "FRK_CfgDef_DeclarationCell"(FieldIndex := 2);
        IF NOT #Image.Rows[#RowIndex].Used OR #Image.Rows[#RowIndex].SchemaVersion <> "FRK_ConfigScratch".Schema
            OR #Image.Rows[#RowIndex].ModelCode <> #Image.Catalog.Codes[#ModelSlot]
            THEN RETURN; END_IF;
        IF NOT "FRK_ConfigRecordValid"(Scope := 'StationB.Satellite.Inner.Cell', Record := #Image.Rows[#RowIndex].Record) THEN RETURN; END_IF;
        #Stored := "FRK_ConfigReserve"(Scope := 'StationB.Satellite.Inner.Cell', Key := 'preset', ModelCode := #Image.Catalog.Codes[#ModelSlot], Reserved := #Targets);
        IF #Stored < 1 OR #Stored > 212 THEN RETURN; END_IF;
        #Targets[#RowIndex] := #Stored;
        #RowIndex := (#ModelSlot - 3) * 26 + 23;
        "FRK_CfgDef_DeclarationCylinder"(FieldIndex := 1);
        IF NOT #Image.Rows[#RowIndex].Used OR #Image.Rows[#RowIndex].SchemaVersion <> "FRK_ConfigScratch".Schema
            OR #Image.Rows[#RowIndex].ModelCode <> #Image.Catalog.Codes[#ModelSlot]
            THEN RETURN; END_IF;
        IF NOT "FRK_ConfigRecordValid"(Scope := 'StationB.Satellite.Inner.Cell.Clamp', Record := #Image.Rows[#RowIndex].Record) THEN RETURN; END_IF;
        #Stored := "FRK_ConfigReserve"(Scope := 'StationB.Satellite.Inner.Cell.Clamp', Key := 'timeout', ModelCode := #Image.Catalog.Codes[#ModelSlot], Reserved := #Targets);
        IF #Stored < 1 OR #Stored > 212 THEN RETURN; END_IF;
        #Targets[#RowIndex] := #Stored;
        #RowIndex := (#ModelSlot - 3) * 26 + 24;
        "FRK_CfgDef_DeclarationCylinder"(FieldIndex := 2);
        IF NOT #Image.Rows[#RowIndex].Used OR #Image.Rows[#RowIndex].SchemaVersion <> "FRK_ConfigScratch".Schema
            OR #Image.Rows[#RowIndex].ModelCode <> #Image.Catalog.Codes[#ModelSlot]
            THEN RETURN; END_IF;
        IF NOT "FRK_ConfigRecordValid"(Scope := 'StationB.Satellite.Inner.Cell.Clamp', Record := #Image.Rows[#RowIndex].Record) THEN RETURN; END_IF;
        #Stored := "FRK_ConfigReserve"(Scope := 'StationB.Satellite.Inner.Cell.Clamp', Key := 'preset', ModelCode := #Image.Catalog.Codes[#ModelSlot], Reserved := #Targets);
        IF #Stored < 1 OR #Stored > 212 THEN RETURN; END_IF;
        #Targets[#RowIndex] := #Stored;
        #RowIndex := (#ModelSlot - 3) * 26 + 25;
        "FRK_CfgDef_DeclarationCylinder"(FieldIndex := 1);
        IF NOT #Image.Rows[#RowIndex].Used OR #Image.Rows[#RowIndex].SchemaVersion <> "FRK_ConfigScratch".Schema
            OR #Image.Rows[#RowIndex].ModelCode <> #Image.Catalog.Codes[#ModelSlot]
            THEN RETURN; END_IF;
        IF NOT "FRK_ConfigRecordValid"(Scope := 'StationB.Satellite.Inner.Cell.Gate', Record := #Image.Rows[#RowIndex].Record) THEN RETURN; END_IF;
        #Stored := "FRK_ConfigReserve"(Scope := 'StationB.Satellite.Inner.Cell.Gate', Key := 'timeout', ModelCode := #Image.Catalog.Codes[#ModelSlot], Reserved := #Targets);
        IF #Stored < 1 OR #Stored > 212 THEN RETURN; END_IF;
        #Targets[#RowIndex] := #Stored;
        #RowIndex := (#ModelSlot - 3) * 26 + 26;
        "FRK_CfgDef_DeclarationCylinder"(FieldIndex := 2);
        IF NOT #Image.Rows[#RowIndex].Used OR #Image.Rows[#RowIndex].SchemaVersion <> "FRK_ConfigScratch".Schema
            OR #Image.Rows[#RowIndex].ModelCode <> #Image.Catalog.Codes[#ModelSlot]
            THEN RETURN; END_IF;
        IF NOT "FRK_ConfigRecordValid"(Scope := 'StationB.Satellite.Inner.Cell.Gate', Record := #Image.Rows[#RowIndex].Record) THEN RETURN; END_IF;
        #Stored := "FRK_ConfigReserve"(Scope := 'StationB.Satellite.Inner.Cell.Gate', Key := 'preset', ModelCode := #Image.Catalog.Codes[#ModelSlot], Reserved := #Targets);
        IF #Stored < 1 OR #Stored > 212 THEN RETURN; END_IF;
        #Targets[#RowIndex] := #Stored;
    END_FOR;
    FOR #Index := 1 TO #Image.RecordCount DO
        "FRK_ConfigStore".Rows[#Targets[#Index]] := #Image.Rows[#Index];
    END_FOR;
    "FRK_ModelStore".Rows[2] := #Image.Catalog;
    "FRK_ConfigStore".SchemaVersion := 1;
    #FRK_ModelApply_R2 := TRUE;
END_FUNCTION
FUNCTION "FRK_ModelCapture" : Bool
{ S7_Optimized_Access := 'TRUE' }
VERSION : 0.1
VAR_INPUT
    RootIndex : Int;
END_VAR
VAR_IN_OUT
    Image : "FRK_ModelImage";
    Catalog : "FRK_ModelCatalog";
END_VAR
BEGIN
    #FRK_ModelCapture := FALSE;
    CASE #RootIndex OF
        1: #FRK_ModelCapture := "FRK_ModelCapture_R1"(Image := #Image, Catalog := #Catalog);
        2: #FRK_ModelCapture := "FRK_ModelCapture_R2"(Image := #Image, Catalog := #Catalog);
        ELSE RETURN;
    END_CASE;
END_FUNCTION
FUNCTION "FRK_ModelApply" : Bool
{ S7_Optimized_Access := 'TRUE' }
VERSION : 0.1
VAR_INPUT
    RootIndex : Int;
END_VAR
VAR_IN_OUT
    Image : "FRK_ModelImage";
END_VAR
BEGIN
    #FRK_ModelApply := FALSE;
    CASE #RootIndex OF
        1: #FRK_ModelApply := "FRK_ModelApply_R1"(Image := #Image);
        2: #FRK_ModelApply := "FRK_ModelApply_R2"(Image := #Image);
        ELSE RETURN;
    END_CASE;
END_FUNCTION
FUNCTION "FRK_ModelDefaults" : Void
{ S7_Optimized_Access := 'TRUE' }
VERSION : 0.1
VAR_INPUT
    RootIndex : Int;
END_VAR
BEGIN
    IF #RootIndex < 1 OR #RootIndex > 2 THEN RETURN; END_IF;
    "FRK_ModelStore".Rows[#RootIndex] := "FRK_ModelRuntime".BlankCatalog;
    "FRK_ModelStore".Rows[#RootIndex].SchemaVersion := 1;
    "FRK_ModelStore".Rows[#RootIndex].Capacity := 3;
    "FRK_ModelStore".Rows[#RootIndex].Count := 2;
    "FRK_ModelStore".Rows[#RootIndex].Generation := 1;
    IF #RootIndex = 1 THEN "FRK_ModelStore".Rows[#RootIndex].Scope := 'StationA'; END_IF;
    IF #RootIndex = 2 THEN "FRK_ModelStore".Rows[#RootIndex].Scope := 'StationB'; END_IF;
    "FRK_ModelStore".Rows[#RootIndex].Codes[1] := 'MODEL_A';
    "FRK_ModelStore".Rows[#RootIndex].Codes[2] := 'MODEL_B';
    "FRK_ModelStore".Rows[#RootIndex].Checksum := "FRK_ModelCrc"(Catalog := "FRK_ModelStore".Rows[#RootIndex]);
END_FUNCTION
FUNCTION "FRK_ModelPrepare" : Void
{ S7_Optimized_Access := 'TRUE' }
VERSION : 0.1
VAR_INPUT
    Startup : Bool;
END_VAR
VAR_TEMP
    RootIndex : Int;
    Index : DInt;
END_VAR
BEGIN
    IF NOT #Startup THEN RETURN; END_IF;
    FOR #RootIndex := 1 TO 2 DO
        "FRK_ModelRuntime".Rows[#RootIndex] := "FRK_ModelRuntime".BlankWork;
    END_FOR;
END_FUNCTION
FUNCTION "FRK_ModelBoot" : Void
{ S7_Optimized_Access := 'TRUE' }
VERSION : 0.1
VAR_INPUT
    Startup : Bool;
END_VAR
VAR_TEMP
    Virgin : Bool;
    Ok : Bool;
END_VAR
BEGIN
    IF NOT #Startup THEN RETURN; END_IF;
    #Virgin := "FRK_ModelVirgin"(Catalog := "FRK_ModelStore".Rows[1]);
    #Ok := "FRK_ModelValid"(RootIndex := 1, Catalog := "FRK_ModelStore".Rows[1]);
    IF #Ok THEN #Ok := "FRK_ModelCapture"(RootIndex := 1, Catalog := "FRK_ModelStore".Rows[1], Image := "FRK_ModelRuntime".ScratchImage); END_IF;
    IF NOT #Ok THEN
        "FRK_ModelDefaults"(RootIndex := 1);
        IF NOT #Virgin THEN "FRK_ConfigLoss"(RootIndex := 1, Scope := 'StationA'); END_IF;
    END_IF;
    IF NOT "FRK_ModelKnown"(RootIndex := 1, Code := "FRK_ConfigStore".ActiveModels[1]) THEN
        "FRK_ConfigSetActiveModel"(RootIndex := 1, ModelCode := 'MODEL_A');
        IF NOT #Virgin OR "FRK_ConfigStore".SchemaVersion <> 0 THEN "FRK_ConfigLoss"(RootIndex := 1, Scope := 'StationA'); END_IF;
    END_IF;
    "FRK_ModelRuntime".Rows[1].Ready := TRUE;
    #Virgin := "FRK_ModelVirgin"(Catalog := "FRK_ModelStore".Rows[2]);
    #Ok := "FRK_ModelValid"(RootIndex := 2, Catalog := "FRK_ModelStore".Rows[2]);
    IF #Ok THEN #Ok := "FRK_ModelCapture"(RootIndex := 2, Catalog := "FRK_ModelStore".Rows[2], Image := "FRK_ModelRuntime".ScratchImage); END_IF;
    IF NOT #Ok THEN
        "FRK_ModelDefaults"(RootIndex := 2);
        IF NOT #Virgin THEN "FRK_ConfigLoss"(RootIndex := 2, Scope := 'StationB'); END_IF;
    END_IF;
    IF NOT "FRK_ModelKnown"(RootIndex := 2, Code := "FRK_ConfigStore".ActiveModels[2]) THEN
        "FRK_ConfigSetActiveModel"(RootIndex := 2, ModelCode := 'MODEL_A');
        IF NOT #Virgin OR "FRK_ConfigStore".SchemaVersion <> 0 THEN "FRK_ConfigLoss"(RootIndex := 2, Scope := 'StationB'); END_IF;
    END_IF;
    "FRK_ModelRuntime".Rows[2].Ready := TRUE;
END_FUNCTION
FUNCTION "FRK_ModelSave" : Void
{ S7_Optimized_Access := 'TRUE' }
VERSION : 0.1
VAR_INPUT
    RootIndex : Int;
END_VAR
BEGIN
    RETURN;
END_FUNCTION
FUNCTION "FRK_ModelSaved" : Bool
{ S7_Optimized_Access := 'TRUE' }
VERSION : 0.1
VAR_INPUT
    RootIndex : Int;
END_VAR
BEGIN
    #FRK_ModelSaved := TRUE;
END_FUNCTION
FUNCTION "FRK_ModelTick" : Bool
{ S7_Optimized_Access := 'TRUE' }
VERSION : 0.1
VAR_INPUT
    RootIndex : Int;
END_VAR
BEGIN
    #FRK_ModelTick := FALSE;
    IF #RootIndex < 1 OR #RootIndex > 2 THEN RETURN; END_IF;
    IF "FRK_ModelRuntime".Rows[#RootIndex].State <> 1 THEN RETURN; END_IF;
    IF NOT "FRK_ModelSaved"(RootIndex := #RootIndex) THEN RETURN; END_IF;
    "FRK_ModelStore".Rows[#RootIndex] := "FRK_ModelRuntime".Rows[#RootIndex].Stage;
    "FRK_ModelRuntime".Rows[#RootIndex].State := 0;
    #FRK_ModelTick := TRUE;
END_FUNCTION
